// TIA Portal V19 export
ORGANIZATION_BLOCK "CyclicInterrupt"   // OB30, LAD, CyclicInterrupt
{ S7_Optimized_Access := 'TRUE' }
// stored: SetENOAutomatically false
   VAR_INPUT
      Initial_Call : Bool;   // Initial call of this OB
      Event_Count : Int;   // Events discarded
   END_VAR
   VAR_TEMP   // added for the SCL form of the ladder/FBD networks
      _w1 : Bool;
      _w2 : Bool;
   END_VAR
BEGIN

REGION Network 1: CHILLED_P01_SPEED_SP
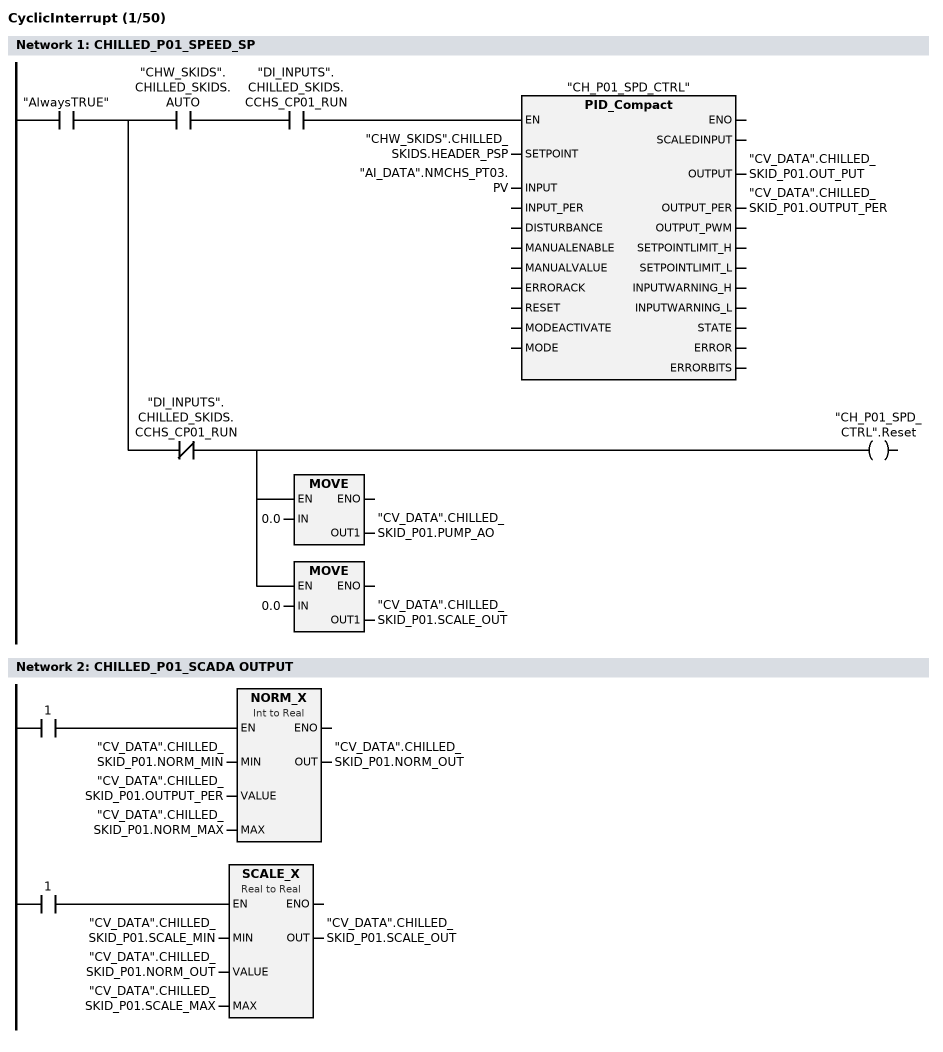
   RUNG wire#powerrail
      Contact( "AlwaysTRUE" )
      wire#w1
      Contact( "CHW_SKIDS".CHILLED_SKIDS.AUTO )
      Contact( "DI_INPUTS".CHILLED_SKIDS.CCHS_CP01_RUN )
      "CH_P01_SPD_CTRL".PID_Compact(Setpoint := "CHW_SKIDS".CHILLED_SKIDS.HEADER_PSP, Input := "AI_DATA".NMCHS_PT03.PV, Input_PER :=, Disturbance :=, ManualEnable :=, ManualValue :=, ErrorAck :=, Reset :=, ModeActivate :=, Mode :=, ScaledInput =>, Output => "CV_DATA".CHILLED_SKID_P01.OUT_PUT, Output_PER => "CV_DATA".CHILLED_SKID_P01.OUTPUT_PER, Output_PWM =>, SetpointLimit_H =>, SetpointLimit_L =>, InputWarning_H =>, InputWarning_L =>, State =>, Error =>, ErrorBits =>)
   END_RUNG
   RUNG wire#w1
      I_Contact( "DI_INPUTS".CHILLED_SKIDS.CCHS_CP01_RUN )
      wire#w2
      Coil( "CH_P01_SPD_CTRL".Reset )
   END_RUNG
   RUNG wire#w2
      Move(in := 0.0, out1 => "CV_DATA".CHILLED_SKID_P01.PUMP_AO)
   END_RUNG
   RUNG wire#w2
      Move(in := 0.0, out1 => "CV_DATA".CHILLED_SKID_P01.SCALE_OUT)
   END_RUNG
   // the same network as SCL:
   #_w1 := "AlwaysTRUE";
   IF "AlwaysTRUE" AND "CHW_SKIDS".CHILLED_SKIDS.AUTO AND "DI_INPUTS".CHILLED_SKIDS.CCHS_CP01_RUN THEN
       "CH_P01_SPD_CTRL"(Setpoint := "CHW_SKIDS".CHILLED_SKIDS.HEADER_PSP,   // PID_Compact
                         Input := "AI_DATA".NMCHS_PT03.PV,
                         Output => "CV_DATA".CHILLED_SKID_P01.OUT_PUT,
                         Output_PER => "CV_DATA".CHILLED_SKID_P01.OUTPUT_PER);
   END_IF;
   "CH_P01_SPD_CTRL".Reset := #_w1 AND NOT "DI_INPUTS".CHILLED_SKIDS.CCHS_CP01_RUN;
   IF "CH_P01_SPD_CTRL".Reset THEN
       "CV_DATA".CHILLED_SKID_P01.PUMP_AO := 0.0;
       "CV_DATA".CHILLED_SKID_P01.SCALE_OUT := 0.0;
   END_IF;
END_REGION

REGION Network 2: CHILLED_P01_SCADA OUTPUT
   RUNG wire#powerrail
      Contact( 1 )
      { S7_Templates := "[SrcType := Int, DestType := Real]" } Normalize(min := "CV_DATA".CHILLED_SKID_P01.NORM_MIN, value := "CV_DATA".CHILLED_SKID_P01.OUTPUT_PER, max := "CV_DATA".CHILLED_SKID_P01.NORM_MAX, out => "CV_DATA".CHILLED_SKID_P01.NORM_OUT)
   END_RUNG
   RUNG wire#powerrail
      Contact( 1 )
      { S7_Templates := "[SrcType := Real, DestType := Real]" } Scale(min := "CV_DATA".CHILLED_SKID_P01.SCALE_MIN, value := "CV_DATA".CHILLED_SKID_P01.NORM_OUT, max := "CV_DATA".CHILLED_SKID_P01.SCALE_MAX, out => "CV_DATA".CHILLED_SKID_P01.SCALE_OUT)
   END_RUNG
   // the same network as SCL:
   IF 1 THEN
       "CV_DATA".CHILLED_SKID_P01.NORM_OUT := NORM_X(MIN := "CV_DATA".CHILLED_SKID_P01.NORM_MIN, VALUE := "CV_DATA".CHILLED_SKID_P01.OUTPUT_PER, MAX := "CV_DATA".CHILLED_SKID_P01.NORM_MAX);
       "CV_DATA".CHILLED_SKID_P01.SCALE_OUT := SCALE_X(MIN := "CV_DATA".CHILLED_SKID_P01.SCALE_MIN, VALUE := "CV_DATA".CHILLED_SKID_P01.NORM_OUT, MAX := "CV_DATA".CHILLED_SKID_P01.SCALE_MAX);
   END_IF;
END_REGION

REGION Network 3: CHILLED_P01_MANUAL OUTPUT
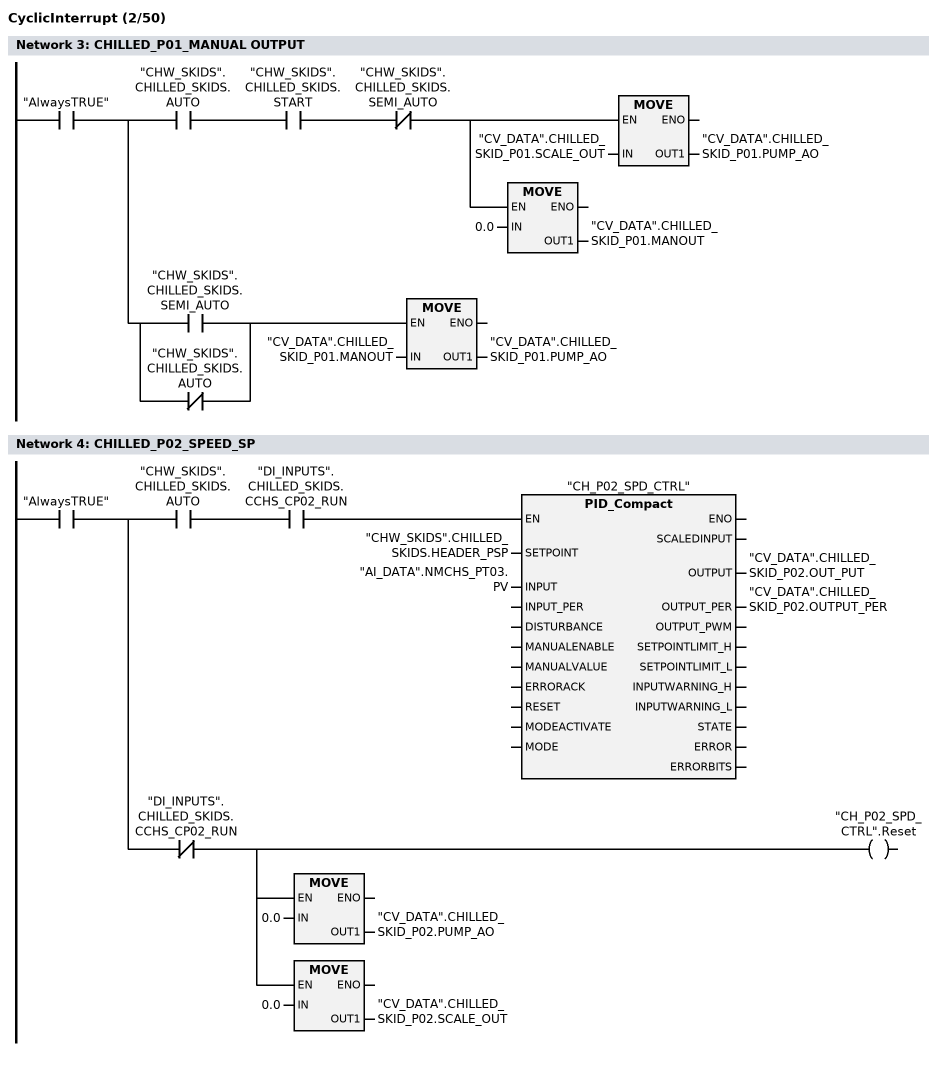
   RUNG wire#powerrail
      Contact( "AlwaysTRUE" )
      wire#w1
      Contact( "CHW_SKIDS".CHILLED_SKIDS.AUTO )
      Contact( "CHW_SKIDS".CHILLED_SKIDS.START )
      I_Contact( "CHW_SKIDS".CHILLED_SKIDS.SEMI_AUTO )
      wire#w2
      Move(in := "CV_DATA".CHILLED_SKID_P01.SCALE_OUT, out1 => "CV_DATA".CHILLED_SKID_P01.PUMP_AO)
   END_RUNG
   RUNG wire#w2
      Move(in := 0.0, out1 => "CV_DATA".CHILLED_SKID_P01.MANOUT)
   END_RUNG
   RUNG wire#w1
      Contact( "CHW_SKIDS".CHILLED_SKIDS.SEMI_AUTO )
      wire#w3
      Move(in := "CV_DATA".CHILLED_SKID_P01.MANOUT, out1 => "CV_DATA".CHILLED_SKID_P01.PUMP_AO)
   END_RUNG
   RUNG wire#w1
      I_Contact( "CHW_SKIDS".CHILLED_SKIDS.AUTO )
   END_RUNG wire#w3
   // the same network as SCL:
   IF "AlwaysTRUE" AND "CHW_SKIDS".CHILLED_SKIDS.AUTO AND "CHW_SKIDS".CHILLED_SKIDS.START AND NOT "CHW_SKIDS".CHILLED_SKIDS.SEMI_AUTO THEN
       "CV_DATA".CHILLED_SKID_P01.PUMP_AO := "CV_DATA".CHILLED_SKID_P01.SCALE_OUT;
       "CV_DATA".CHILLED_SKID_P01.MANOUT := 0.0;
   END_IF;
   IF "AlwaysTRUE" AND ("CHW_SKIDS".CHILLED_SKIDS.SEMI_AUTO OR NOT "CHW_SKIDS".CHILLED_SKIDS.AUTO) THEN
       "CV_DATA".CHILLED_SKID_P01.PUMP_AO := "CV_DATA".CHILLED_SKID_P01.MANOUT;
   END_IF;
END_REGION

REGION Network 4: CHILLED_P02_SPEED_SP
   RUNG wire#powerrail
      Contact( "AlwaysTRUE" )
      wire#w1
      Contact( "CHW_SKIDS".CHILLED_SKIDS.AUTO )
      Contact( "DI_INPUTS".CHILLED_SKIDS.CCHS_CP02_RUN )
      "CH_P02_SPD_CTRL".PID_Compact(Setpoint := "CHW_SKIDS".CHILLED_SKIDS.HEADER_PSP, Input := "AI_DATA".NMCHS_PT03.PV, Input_PER :=, Disturbance :=, ManualEnable :=, ManualValue :=, ErrorAck :=, Reset :=, ModeActivate :=, Mode :=, ScaledInput =>, Output => "CV_DATA".CHILLED_SKID_P02.OUT_PUT, Output_PER => "CV_DATA".CHILLED_SKID_P02.OUTPUT_PER, Output_PWM =>, SetpointLimit_H =>, SetpointLimit_L =>, InputWarning_H =>, InputWarning_L =>, State =>, Error =>, ErrorBits =>)
   END_RUNG
   RUNG wire#w1
      I_Contact( "DI_INPUTS".CHILLED_SKIDS.CCHS_CP02_RUN )
      wire#w2
      Coil( "CH_P02_SPD_CTRL".Reset )
   END_RUNG
   RUNG wire#w2
      Move(in := 0.0, out1 => "CV_DATA".CHILLED_SKID_P02.PUMP_AO)
   END_RUNG
   RUNG wire#w2
      Move(in := 0.0, out1 => "CV_DATA".CHILLED_SKID_P02.SCALE_OUT)
   END_RUNG
   // the same network as SCL:
   #_w1 := "AlwaysTRUE";
   IF "AlwaysTRUE" AND "CHW_SKIDS".CHILLED_SKIDS.AUTO AND "DI_INPUTS".CHILLED_SKIDS.CCHS_CP02_RUN THEN
       "CH_P02_SPD_CTRL"(Setpoint := "CHW_SKIDS".CHILLED_SKIDS.HEADER_PSP,   // PID_Compact
                         Input := "AI_DATA".NMCHS_PT03.PV,
                         Output => "CV_DATA".CHILLED_SKID_P02.OUT_PUT,
                         Output_PER => "CV_DATA".CHILLED_SKID_P02.OUTPUT_PER);
   END_IF;
   "CH_P02_SPD_CTRL".Reset := #_w1 AND NOT "DI_INPUTS".CHILLED_SKIDS.CCHS_CP02_RUN;
   IF "CH_P02_SPD_CTRL".Reset THEN
       "CV_DATA".CHILLED_SKID_P02.PUMP_AO := 0.0;
       "CV_DATA".CHILLED_SKID_P02.SCALE_OUT := 0.0;
   END_IF;
END_REGION

REGION Network 5: CHILLED_P02_SCADA OUTPUT
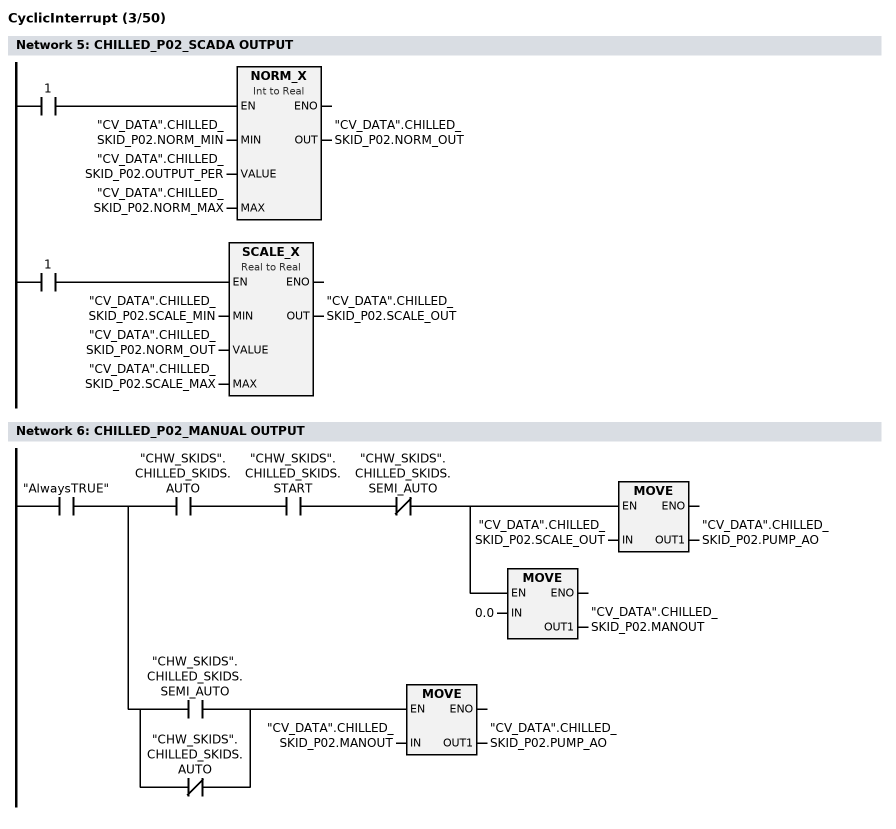
   RUNG wire#powerrail
      Contact( 1 )
      { S7_Templates := "[SrcType := Int, DestType := Real]" } Normalize(min := "CV_DATA".CHILLED_SKID_P02.NORM_MIN, value := "CV_DATA".CHILLED_SKID_P02.OUTPUT_PER, max := "CV_DATA".CHILLED_SKID_P02.NORM_MAX, out => "CV_DATA".CHILLED_SKID_P02.NORM_OUT)
   END_RUNG
   RUNG wire#powerrail
      Contact( 1 )
      { S7_Templates := "[SrcType := Real, DestType := Real]" } Scale(min := "CV_DATA".CHILLED_SKID_P02.SCALE_MIN, value := "CV_DATA".CHILLED_SKID_P02.NORM_OUT, max := "CV_DATA".CHILLED_SKID_P02.SCALE_MAX, out => "CV_DATA".CHILLED_SKID_P02.SCALE_OUT)
   END_RUNG
   // the same network as SCL:
   IF 1 THEN
       "CV_DATA".CHILLED_SKID_P02.NORM_OUT := NORM_X(MIN := "CV_DATA".CHILLED_SKID_P02.NORM_MIN, VALUE := "CV_DATA".CHILLED_SKID_P02.OUTPUT_PER, MAX := "CV_DATA".CHILLED_SKID_P02.NORM_MAX);
       "CV_DATA".CHILLED_SKID_P02.SCALE_OUT := SCALE_X(MIN := "CV_DATA".CHILLED_SKID_P02.SCALE_MIN, VALUE := "CV_DATA".CHILLED_SKID_P02.NORM_OUT, MAX := "CV_DATA".CHILLED_SKID_P02.SCALE_MAX);
   END_IF;
END_REGION

REGION Network 6: CHILLED_P02_MANUAL OUTPUT
   RUNG wire#powerrail
      Contact( "AlwaysTRUE" )
      wire#w1
      Contact( "CHW_SKIDS".CHILLED_SKIDS.AUTO )
      Contact( "CHW_SKIDS".CHILLED_SKIDS.START )
      I_Contact( "CHW_SKIDS".CHILLED_SKIDS.SEMI_AUTO )
      wire#w2
      Move(in := "CV_DATA".CHILLED_SKID_P02.SCALE_OUT, out1 => "CV_DATA".CHILLED_SKID_P02.PUMP_AO)
   END_RUNG
   RUNG wire#w2
      Move(in := 0.0, out1 => "CV_DATA".CHILLED_SKID_P02.MANOUT)
   END_RUNG
   RUNG wire#w1
      Contact( "CHW_SKIDS".CHILLED_SKIDS.SEMI_AUTO )
      wire#w3
      Move(in := "CV_DATA".CHILLED_SKID_P02.MANOUT, out1 => "CV_DATA".CHILLED_SKID_P02.PUMP_AO)
   END_RUNG
   RUNG wire#w1
      I_Contact( "CHW_SKIDS".CHILLED_SKIDS.AUTO )
   END_RUNG wire#w3
   // the same network as SCL:
   IF "AlwaysTRUE" AND "CHW_SKIDS".CHILLED_SKIDS.AUTO AND "CHW_SKIDS".CHILLED_SKIDS.START AND NOT "CHW_SKIDS".CHILLED_SKIDS.SEMI_AUTO THEN
       "CV_DATA".CHILLED_SKID_P02.PUMP_AO := "CV_DATA".CHILLED_SKID_P02.SCALE_OUT;
       "CV_DATA".CHILLED_SKID_P02.MANOUT := 0.0;
   END_IF;
   IF "AlwaysTRUE" AND ("CHW_SKIDS".CHILLED_SKIDS.SEMI_AUTO OR NOT "CHW_SKIDS".CHILLED_SKIDS.AUTO) THEN
       "CV_DATA".CHILLED_SKID_P02.PUMP_AO := "CV_DATA".CHILLED_SKID_P02.MANOUT;
   END_IF;
END_REGION

REGION Network 7: CHILLED_P03_SPEED_SP
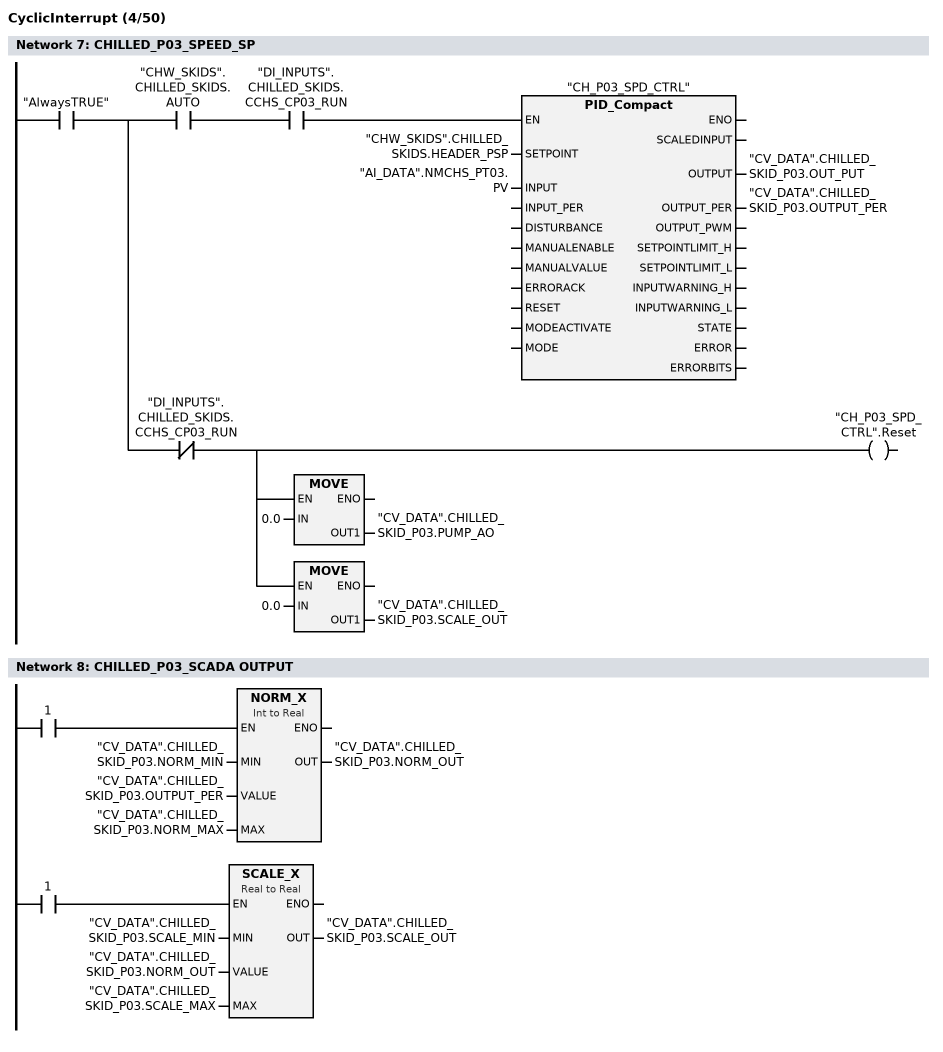
   RUNG wire#powerrail
      Contact( "AlwaysTRUE" )
      wire#w1
      Contact( "CHW_SKIDS".CHILLED_SKIDS.AUTO )
      Contact( "DI_INPUTS".CHILLED_SKIDS.CCHS_CP03_RUN )
      "CH_P03_SPD_CTRL".PID_Compact(Setpoint := "CHW_SKIDS".CHILLED_SKIDS.HEADER_PSP, Input := "AI_DATA".NMCHS_PT03.PV, Input_PER :=, Disturbance :=, ManualEnable :=, ManualValue :=, ErrorAck :=, Reset :=, ModeActivate :=, Mode :=, ScaledInput =>, Output => "CV_DATA".CHILLED_SKID_P03.OUT_PUT, Output_PER => "CV_DATA".CHILLED_SKID_P03.OUTPUT_PER, Output_PWM =>, SetpointLimit_H =>, SetpointLimit_L =>, InputWarning_H =>, InputWarning_L =>, State =>, Error =>, ErrorBits =>)
   END_RUNG
   RUNG wire#w1
      I_Contact( "DI_INPUTS".CHILLED_SKIDS.CCHS_CP03_RUN )
      wire#w2
      Coil( "CH_P03_SPD_CTRL".Reset )
   END_RUNG
   RUNG wire#w2
      Move(in := 0.0, out1 => "CV_DATA".CHILLED_SKID_P03.PUMP_AO)
   END_RUNG
   RUNG wire#w2
      Move(in := 0.0, out1 => "CV_DATA".CHILLED_SKID_P03.SCALE_OUT)
   END_RUNG
   // the same network as SCL:
   #_w1 := "AlwaysTRUE";
   IF "AlwaysTRUE" AND "CHW_SKIDS".CHILLED_SKIDS.AUTO AND "DI_INPUTS".CHILLED_SKIDS.CCHS_CP03_RUN THEN
       "CH_P03_SPD_CTRL"(Setpoint := "CHW_SKIDS".CHILLED_SKIDS.HEADER_PSP,   // PID_Compact
                         Input := "AI_DATA".NMCHS_PT03.PV,
                         Output => "CV_DATA".CHILLED_SKID_P03.OUT_PUT,
                         Output_PER => "CV_DATA".CHILLED_SKID_P03.OUTPUT_PER);
   END_IF;
   "CH_P03_SPD_CTRL".Reset := #_w1 AND NOT "DI_INPUTS".CHILLED_SKIDS.CCHS_CP03_RUN;
   IF "CH_P03_SPD_CTRL".Reset THEN
       "CV_DATA".CHILLED_SKID_P03.PUMP_AO := 0.0;
       "CV_DATA".CHILLED_SKID_P03.SCALE_OUT := 0.0;
   END_IF;
END_REGION

REGION Network 8: CHILLED_P03_SCADA OUTPUT
   RUNG wire#powerrail
      Contact( 1 )
      { S7_Templates := "[SrcType := Int, DestType := Real]" } Normalize(min := "CV_DATA".CHILLED_SKID_P03.NORM_MIN, value := "CV_DATA".CHILLED_SKID_P03.OUTPUT_PER, max := "CV_DATA".CHILLED_SKID_P03.NORM_MAX, out => "CV_DATA".CHILLED_SKID_P03.NORM_OUT)
   END_RUNG
   RUNG wire#powerrail
      Contact( 1 )
      { S7_Templates := "[SrcType := Real, DestType := Real]" } Scale(min := "CV_DATA".CHILLED_SKID_P03.SCALE_MIN, value := "CV_DATA".CHILLED_SKID_P03.NORM_OUT, max := "CV_DATA".CHILLED_SKID_P03.SCALE_MAX, out => "CV_DATA".CHILLED_SKID_P03.SCALE_OUT)
   END_RUNG
   // the same network as SCL:
   IF 1 THEN
       "CV_DATA".CHILLED_SKID_P03.NORM_OUT := NORM_X(MIN := "CV_DATA".CHILLED_SKID_P03.NORM_MIN, VALUE := "CV_DATA".CHILLED_SKID_P03.OUTPUT_PER, MAX := "CV_DATA".CHILLED_SKID_P03.NORM_MAX);
       "CV_DATA".CHILLED_SKID_P03.SCALE_OUT := SCALE_X(MIN := "CV_DATA".CHILLED_SKID_P03.SCALE_MIN, VALUE := "CV_DATA".CHILLED_SKID_P03.NORM_OUT, MAX := "CV_DATA".CHILLED_SKID_P03.SCALE_MAX);
   END_IF;
END_REGION

REGION Network 9: CHILLED_P03_MANUAL OUTPUT
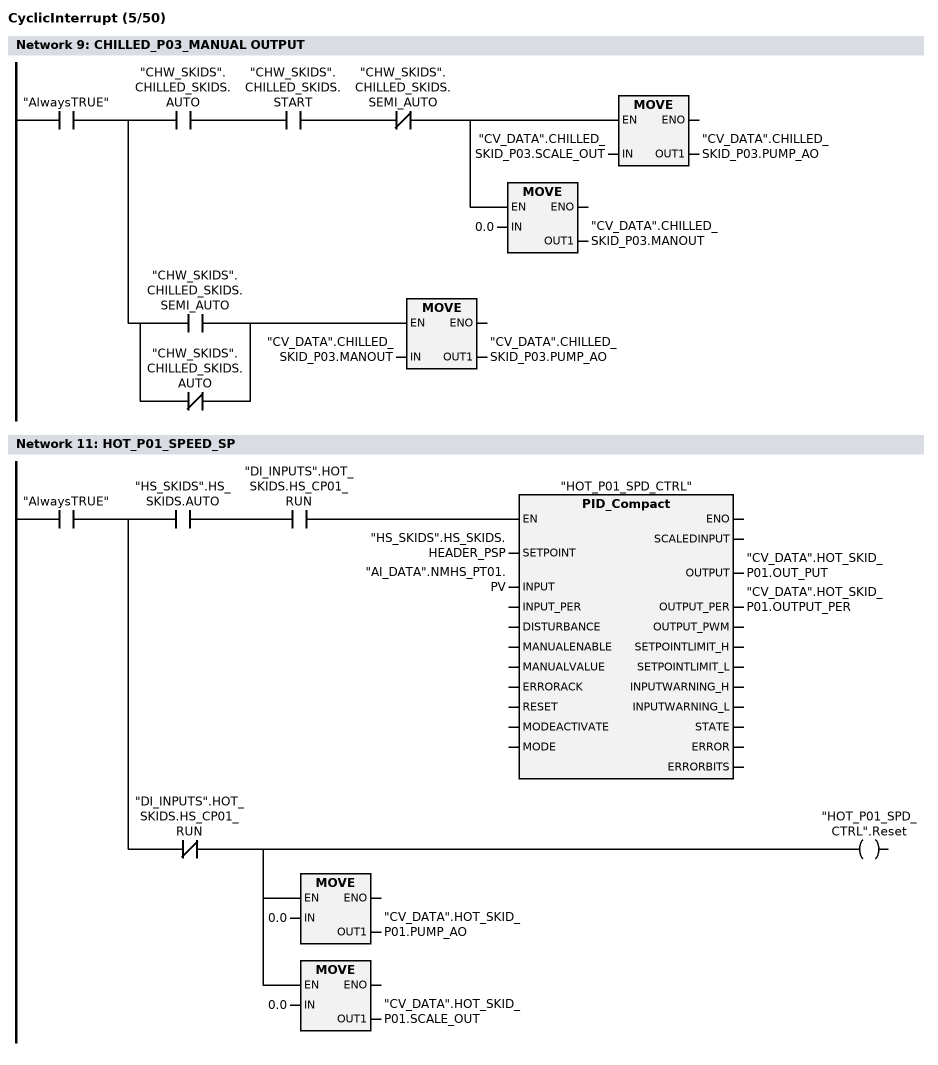
   RUNG wire#powerrail
      Contact( "AlwaysTRUE" )
      wire#w1
      Contact( "CHW_SKIDS".CHILLED_SKIDS.AUTO )
      Contact( "CHW_SKIDS".CHILLED_SKIDS.START )
      I_Contact( "CHW_SKIDS".CHILLED_SKIDS.SEMI_AUTO )
      wire#w2
      Move(in := "CV_DATA".CHILLED_SKID_P03.SCALE_OUT, out1 => "CV_DATA".CHILLED_SKID_P03.PUMP_AO)
   END_RUNG
   RUNG wire#w2
      Move(in := 0.0, out1 => "CV_DATA".CHILLED_SKID_P03.MANOUT)
   END_RUNG
   RUNG wire#w1
      Contact( "CHW_SKIDS".CHILLED_SKIDS.SEMI_AUTO )
      wire#w3
      Move(in := "CV_DATA".CHILLED_SKID_P03.MANOUT, out1 => "CV_DATA".CHILLED_SKID_P03.PUMP_AO)
   END_RUNG
   RUNG wire#w1
      I_Contact( "CHW_SKIDS".CHILLED_SKIDS.AUTO )
   END_RUNG wire#w3
   // the same network as SCL:
   IF "AlwaysTRUE" AND "CHW_SKIDS".CHILLED_SKIDS.AUTO AND "CHW_SKIDS".CHILLED_SKIDS.START AND NOT "CHW_SKIDS".CHILLED_SKIDS.SEMI_AUTO THEN
       "CV_DATA".CHILLED_SKID_P03.PUMP_AO := "CV_DATA".CHILLED_SKID_P03.SCALE_OUT;
       "CV_DATA".CHILLED_SKID_P03.MANOUT := 0.0;
   END_IF;
   IF "AlwaysTRUE" AND ("CHW_SKIDS".CHILLED_SKIDS.SEMI_AUTO OR NOT "CHW_SKIDS".CHILLED_SKIDS.AUTO) THEN
       "CV_DATA".CHILLED_SKID_P03.PUMP_AO := "CV_DATA".CHILLED_SKID_P03.MANOUT;
   END_IF;
END_REGION

REGION Network 11: HOT_P01_SPEED_SP
   RUNG wire#powerrail
      Contact( "AlwaysTRUE" )
      wire#w1
      Contact( "HS_SKIDS".HS_SKIDS.AUTO )
      Contact( "DI_INPUTS".HOT_SKIDS.HS_CP01_RUN )
      "HOT_P01_SPD_CTRL".PID_Compact(Setpoint := "HS_SKIDS".HS_SKIDS.HEADER_PSP, Input := "AI_DATA".NMHS_PT01.PV, Input_PER :=, Disturbance :=, ManualEnable :=, ManualValue :=, ErrorAck :=, Reset :=, ModeActivate :=, Mode :=, ScaledInput =>, Output => "CV_DATA".HOT_SKID_P01.OUT_PUT, Output_PER => "CV_DATA".HOT_SKID_P01.OUTPUT_PER, Output_PWM =>, SetpointLimit_H =>, SetpointLimit_L =>, InputWarning_H =>, InputWarning_L =>, State =>, Error =>, ErrorBits =>)
   END_RUNG
   RUNG wire#w1
      I_Contact( "DI_INPUTS".HOT_SKIDS.HS_CP01_RUN )
      wire#w2
      Coil( "HOT_P01_SPD_CTRL".Reset )
   END_RUNG
   RUNG wire#w2
      Move(in := 0.0, out1 => "CV_DATA".HOT_SKID_P01.PUMP_AO)
   END_RUNG
   RUNG wire#w2
      Move(in := 0.0, out1 => "CV_DATA".HOT_SKID_P01.SCALE_OUT)
   END_RUNG
   // the same network as SCL:
   #_w1 := "AlwaysTRUE";
   IF "AlwaysTRUE" AND "HS_SKIDS".HS_SKIDS.AUTO AND "DI_INPUTS".HOT_SKIDS.HS_CP01_RUN THEN
       "HOT_P01_SPD_CTRL"(Setpoint := "HS_SKIDS".HS_SKIDS.HEADER_PSP,   // PID_Compact
                          Input := "AI_DATA".NMHS_PT01.PV,
                          Output => "CV_DATA".HOT_SKID_P01.OUT_PUT,
                          Output_PER => "CV_DATA".HOT_SKID_P01.OUTPUT_PER);
   END_IF;
   "HOT_P01_SPD_CTRL".Reset := #_w1 AND NOT "DI_INPUTS".HOT_SKIDS.HS_CP01_RUN;
   IF "HOT_P01_SPD_CTRL".Reset THEN
       "CV_DATA".HOT_SKID_P01.PUMP_AO := 0.0;
       "CV_DATA".HOT_SKID_P01.SCALE_OUT := 0.0;
   END_IF;
END_REGION

REGION Network 12: HOT_P01_SCADA OUTPUT
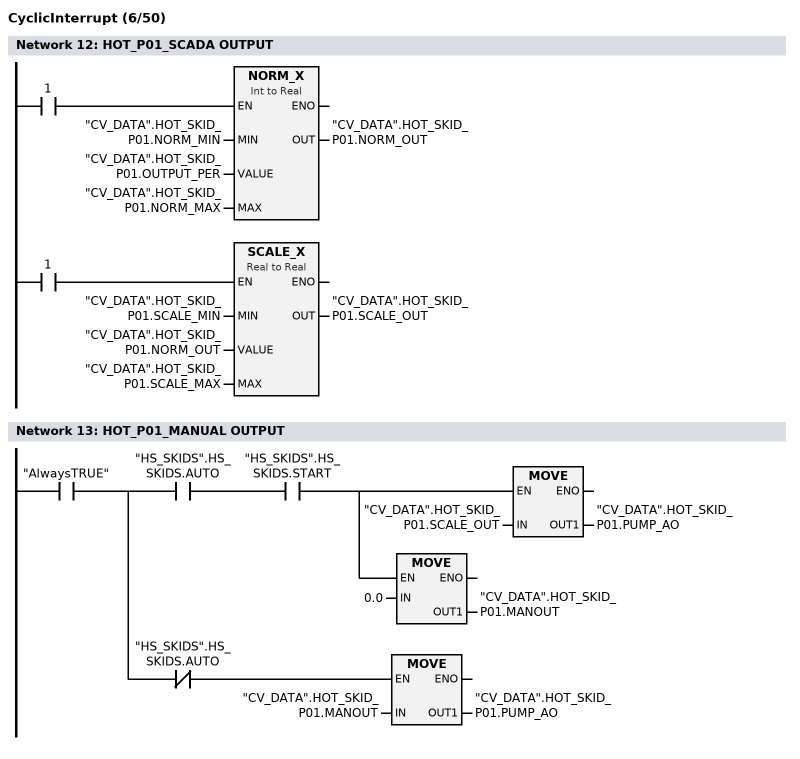
   RUNG wire#powerrail
      Contact( 1 )
      { S7_Templates := "[SrcType := Int, DestType := Real]" } Normalize(min := "CV_DATA".HOT_SKID_P01.NORM_MIN, value := "CV_DATA".HOT_SKID_P01.OUTPUT_PER, max := "CV_DATA".HOT_SKID_P01.NORM_MAX, out => "CV_DATA".HOT_SKID_P01.NORM_OUT)
   END_RUNG
   RUNG wire#powerrail
      Contact( 1 )
      { S7_Templates := "[SrcType := Real, DestType := Real]" } Scale(min := "CV_DATA".HOT_SKID_P01.SCALE_MIN, value := "CV_DATA".HOT_SKID_P01.NORM_OUT, max := "CV_DATA".HOT_SKID_P01.SCALE_MAX, out => "CV_DATA".HOT_SKID_P01.SCALE_OUT)
   END_RUNG
   // the same network as SCL:
   IF 1 THEN
       "CV_DATA".HOT_SKID_P01.NORM_OUT := NORM_X(MIN := "CV_DATA".HOT_SKID_P01.NORM_MIN, VALUE := "CV_DATA".HOT_SKID_P01.OUTPUT_PER, MAX := "CV_DATA".HOT_SKID_P01.NORM_MAX);
       "CV_DATA".HOT_SKID_P01.SCALE_OUT := SCALE_X(MIN := "CV_DATA".HOT_SKID_P01.SCALE_MIN, VALUE := "CV_DATA".HOT_SKID_P01.NORM_OUT, MAX := "CV_DATA".HOT_SKID_P01.SCALE_MAX);
   END_IF;
END_REGION

REGION Network 13: HOT_P01_MANUAL OUTPUT
   RUNG wire#powerrail
      Contact( "AlwaysTRUE" )
      wire#w1
      Contact( "HS_SKIDS".HS_SKIDS.AUTO )
      Contact( "HS_SKIDS".HS_SKIDS.START )
      wire#w2
      Move(in := "CV_DATA".HOT_SKID_P01.SCALE_OUT, out1 => "CV_DATA".HOT_SKID_P01.PUMP_AO)
   END_RUNG
   RUNG wire#w2
      Move(in := 0.0, out1 => "CV_DATA".HOT_SKID_P01.MANOUT)
   END_RUNG
   RUNG wire#w1
      I_Contact( "HS_SKIDS".HS_SKIDS.AUTO )
      Move(in := "CV_DATA".HOT_SKID_P01.MANOUT, out1 => "CV_DATA".HOT_SKID_P01.PUMP_AO)
   END_RUNG
   // the same network as SCL:
   IF "AlwaysTRUE" AND "HS_SKIDS".HS_SKIDS.AUTO AND "HS_SKIDS".HS_SKIDS.START THEN
       "CV_DATA".HOT_SKID_P01.PUMP_AO := "CV_DATA".HOT_SKID_P01.SCALE_OUT;
       "CV_DATA".HOT_SKID_P01.MANOUT := 0.0;
   END_IF;
   IF "AlwaysTRUE" AND NOT "HS_SKIDS".HS_SKIDS.AUTO THEN
       "CV_DATA".HOT_SKID_P01.PUMP_AO := "CV_DATA".HOT_SKID_P01.MANOUT;
   END_IF;
END_REGION

REGION Network 14: HOT_P02_SPEED_SP
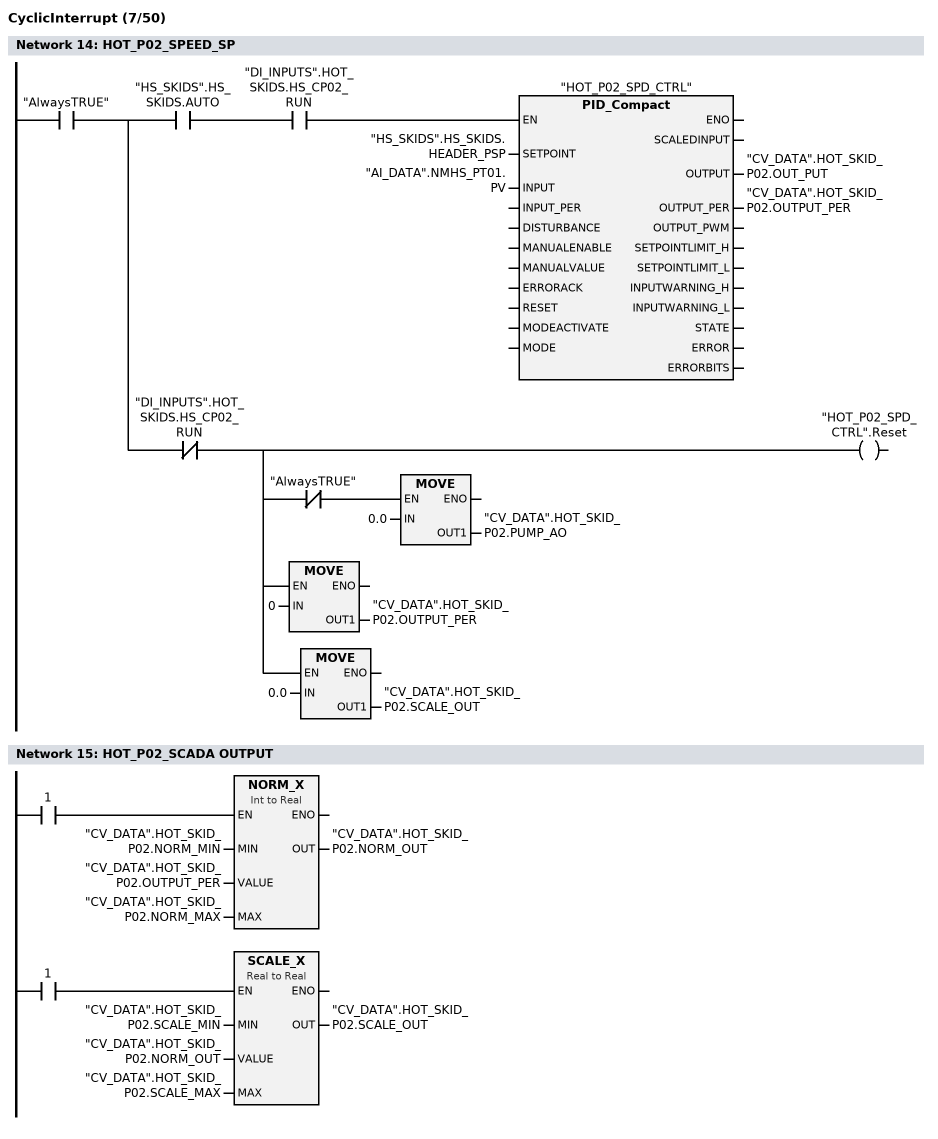
   RUNG wire#powerrail
      Contact( "AlwaysTRUE" )
      wire#w1
      Contact( "HS_SKIDS".HS_SKIDS.AUTO )
      Contact( "DI_INPUTS".HOT_SKIDS.HS_CP02_RUN )
      "HOT_P02_SPD_CTRL".PID_Compact(Setpoint := "HS_SKIDS".HS_SKIDS.HEADER_PSP, Input := "AI_DATA".NMHS_PT01.PV, Input_PER :=, Disturbance :=, ManualEnable :=, ManualValue :=, ErrorAck :=, Reset :=, ModeActivate :=, Mode :=, ScaledInput =>, Output => "CV_DATA".HOT_SKID_P02.OUT_PUT, Output_PER => "CV_DATA".HOT_SKID_P02.OUTPUT_PER, Output_PWM =>, SetpointLimit_H =>, SetpointLimit_L =>, InputWarning_H =>, InputWarning_L =>, State =>, Error =>, ErrorBits =>)
   END_RUNG
   RUNG wire#w1
      I_Contact( "DI_INPUTS".HOT_SKIDS.HS_CP02_RUN )
      wire#w2
      Coil( "HOT_P02_SPD_CTRL".Reset )
   END_RUNG
   RUNG wire#w2
      I_Contact( "AlwaysTRUE" )
      Move(in := 0.0, out1 => "CV_DATA".HOT_SKID_P02.PUMP_AO)
   END_RUNG
   RUNG wire#w2
      Move(in := 0, out1 => "CV_DATA".HOT_SKID_P02.OUTPUT_PER)
   END_RUNG
   RUNG wire#w2
      Move(in := 0.0, out1 => "CV_DATA".HOT_SKID_P02.SCALE_OUT)
   END_RUNG
   // the same network as SCL:
   #_w1 := "AlwaysTRUE";
   IF "AlwaysTRUE" AND "HS_SKIDS".HS_SKIDS.AUTO AND "DI_INPUTS".HOT_SKIDS.HS_CP02_RUN THEN
       "HOT_P02_SPD_CTRL"(Setpoint := "HS_SKIDS".HS_SKIDS.HEADER_PSP,   // PID_Compact
                          Input := "AI_DATA".NMHS_PT01.PV,
                          Output => "CV_DATA".HOT_SKID_P02.OUT_PUT,
                          Output_PER => "CV_DATA".HOT_SKID_P02.OUTPUT_PER);
   END_IF;
   "HOT_P02_SPD_CTRL".Reset := #_w1 AND NOT "DI_INPUTS".HOT_SKIDS.HS_CP02_RUN;
   IF "HOT_P02_SPD_CTRL".Reset AND NOT "AlwaysTRUE" THEN "CV_DATA".HOT_SKID_P02.PUMP_AO := 0.0; END_IF;
   IF "HOT_P02_SPD_CTRL".Reset THEN
       "CV_DATA".HOT_SKID_P02.OUTPUT_PER := 0;
       "CV_DATA".HOT_SKID_P02.SCALE_OUT := 0.0;
   END_IF;
END_REGION

REGION Network 15: HOT_P02_SCADA OUTPUT
   RUNG wire#powerrail
      Contact( 1 )
      { S7_Templates := "[SrcType := Int, DestType := Real]" } Normalize(min := "CV_DATA".HOT_SKID_P02.NORM_MIN, value := "CV_DATA".HOT_SKID_P02.OUTPUT_PER, max := "CV_DATA".HOT_SKID_P02.NORM_MAX, out => "CV_DATA".HOT_SKID_P02.NORM_OUT)
   END_RUNG
   RUNG wire#powerrail
      Contact( 1 )
      { S7_Templates := "[SrcType := Real, DestType := Real]" } Scale(min := "CV_DATA".HOT_SKID_P02.SCALE_MIN, value := "CV_DATA".HOT_SKID_P02.NORM_OUT, max := "CV_DATA".HOT_SKID_P02.SCALE_MAX, out => "CV_DATA".HOT_SKID_P02.SCALE_OUT)
   END_RUNG
   // the same network as SCL:
   IF 1 THEN
       "CV_DATA".HOT_SKID_P02.NORM_OUT := NORM_X(MIN := "CV_DATA".HOT_SKID_P02.NORM_MIN, VALUE := "CV_DATA".HOT_SKID_P02.OUTPUT_PER, MAX := "CV_DATA".HOT_SKID_P02.NORM_MAX);
       "CV_DATA".HOT_SKID_P02.SCALE_OUT := SCALE_X(MIN := "CV_DATA".HOT_SKID_P02.SCALE_MIN, VALUE := "CV_DATA".HOT_SKID_P02.NORM_OUT, MAX := "CV_DATA".HOT_SKID_P02.SCALE_MAX);
   END_IF;
END_REGION

REGION Network 16: HOT_P02_MANUAL OUTPUT
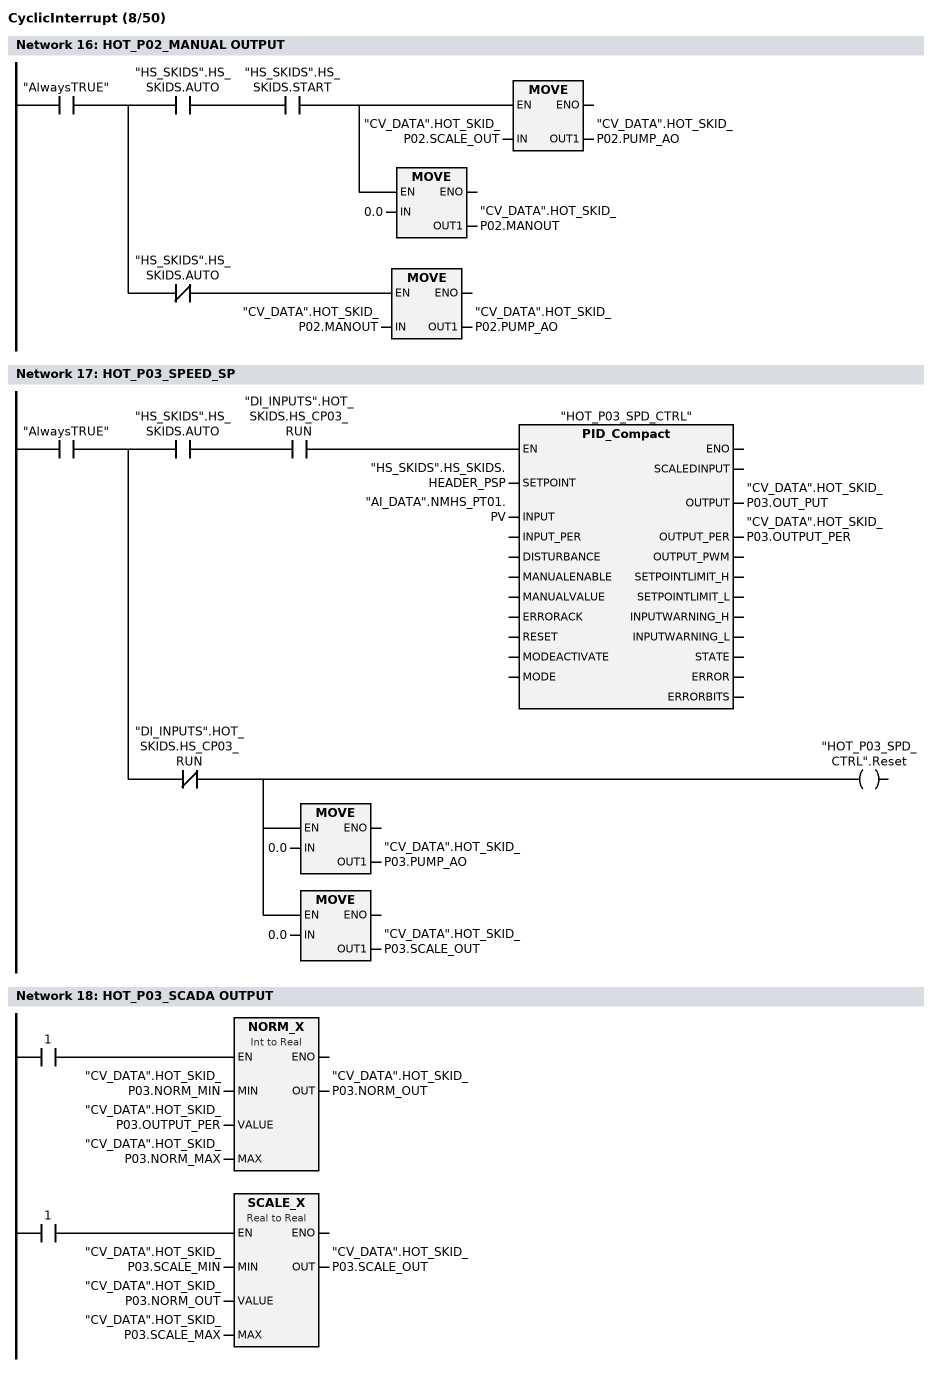
   RUNG wire#powerrail
      Contact( "AlwaysTRUE" )
      wire#w1
      Contact( "HS_SKIDS".HS_SKIDS.AUTO )
      Contact( "HS_SKIDS".HS_SKIDS.START )
      wire#w2
      Move(in := "CV_DATA".HOT_SKID_P02.SCALE_OUT, out1 => "CV_DATA".HOT_SKID_P02.PUMP_AO)
   END_RUNG
   RUNG wire#w2
      Move(in := 0.0, out1 => "CV_DATA".HOT_SKID_P02.MANOUT)
   END_RUNG
   RUNG wire#w1
      I_Contact( "HS_SKIDS".HS_SKIDS.AUTO )
      Move(in := "CV_DATA".HOT_SKID_P02.MANOUT, out1 => "CV_DATA".HOT_SKID_P02.PUMP_AO)
   END_RUNG
   // the same network as SCL:
   IF "AlwaysTRUE" AND "HS_SKIDS".HS_SKIDS.AUTO AND "HS_SKIDS".HS_SKIDS.START THEN
       "CV_DATA".HOT_SKID_P02.PUMP_AO := "CV_DATA".HOT_SKID_P02.SCALE_OUT;
       "CV_DATA".HOT_SKID_P02.MANOUT := 0.0;
   END_IF;
   IF "AlwaysTRUE" AND NOT "HS_SKIDS".HS_SKIDS.AUTO THEN
       "CV_DATA".HOT_SKID_P02.PUMP_AO := "CV_DATA".HOT_SKID_P02.MANOUT;
   END_IF;
END_REGION

REGION Network 17: HOT_P03_SPEED_SP
   RUNG wire#powerrail
      Contact( "AlwaysTRUE" )
      wire#w1
      Contact( "HS_SKIDS".HS_SKIDS.AUTO )
      Contact( "DI_INPUTS".HOT_SKIDS.HS_CP03_RUN )
      "HOT_P03_SPD_CTRL".PID_Compact(Setpoint := "HS_SKIDS".HS_SKIDS.HEADER_PSP, Input := "AI_DATA".NMHS_PT01.PV, Input_PER :=, Disturbance :=, ManualEnable :=, ManualValue :=, ErrorAck :=, Reset :=, ModeActivate :=, Mode :=, ScaledInput =>, Output => "CV_DATA".HOT_SKID_P03.OUT_PUT, Output_PER => "CV_DATA".HOT_SKID_P03.OUTPUT_PER, Output_PWM =>, SetpointLimit_H =>, SetpointLimit_L =>, InputWarning_H =>, InputWarning_L =>, State =>, Error =>, ErrorBits =>)
   END_RUNG
   RUNG wire#w1
      I_Contact( "DI_INPUTS".HOT_SKIDS.HS_CP03_RUN )
      wire#w2
      Coil( "HOT_P03_SPD_CTRL".Reset )
   END_RUNG
   RUNG wire#w2
      Move(in := 0.0, out1 => "CV_DATA".HOT_SKID_P03.PUMP_AO)
   END_RUNG
   RUNG wire#w2
      Move(in := 0.0, out1 => "CV_DATA".HOT_SKID_P03.SCALE_OUT)
   END_RUNG
   // the same network as SCL:
   #_w1 := "AlwaysTRUE";
   IF "AlwaysTRUE" AND "HS_SKIDS".HS_SKIDS.AUTO AND "DI_INPUTS".HOT_SKIDS.HS_CP03_RUN THEN
       "HOT_P03_SPD_CTRL"(Setpoint := "HS_SKIDS".HS_SKIDS.HEADER_PSP,   // PID_Compact
                          Input := "AI_DATA".NMHS_PT01.PV,
                          Output => "CV_DATA".HOT_SKID_P03.OUT_PUT,
                          Output_PER => "CV_DATA".HOT_SKID_P03.OUTPUT_PER);
   END_IF;
   "HOT_P03_SPD_CTRL".Reset := #_w1 AND NOT "DI_INPUTS".HOT_SKIDS.HS_CP03_RUN;
   IF "HOT_P03_SPD_CTRL".Reset THEN
       "CV_DATA".HOT_SKID_P03.PUMP_AO := 0.0;
       "CV_DATA".HOT_SKID_P03.SCALE_OUT := 0.0;
   END_IF;
END_REGION

REGION Network 18: HOT_P03_SCADA OUTPUT
   RUNG wire#powerrail
      Contact( 1 )
      { S7_Templates := "[SrcType := Int, DestType := Real]" } Normalize(min := "CV_DATA".HOT_SKID_P03.NORM_MIN, value := "CV_DATA".HOT_SKID_P03.OUTPUT_PER, max := "CV_DATA".HOT_SKID_P03.NORM_MAX, out => "CV_DATA".HOT_SKID_P03.NORM_OUT)
   END_RUNG
   RUNG wire#powerrail
      Contact( 1 )
      { S7_Templates := "[SrcType := Real, DestType := Real]" } Scale(min := "CV_DATA".HOT_SKID_P03.SCALE_MIN, value := "CV_DATA".HOT_SKID_P03.NORM_OUT, max := "CV_DATA".HOT_SKID_P03.SCALE_MAX, out => "CV_DATA".HOT_SKID_P03.SCALE_OUT)
   END_RUNG
   // the same network as SCL:
   IF 1 THEN
       "CV_DATA".HOT_SKID_P03.NORM_OUT := NORM_X(MIN := "CV_DATA".HOT_SKID_P03.NORM_MIN, VALUE := "CV_DATA".HOT_SKID_P03.OUTPUT_PER, MAX := "CV_DATA".HOT_SKID_P03.NORM_MAX);
       "CV_DATA".HOT_SKID_P03.SCALE_OUT := SCALE_X(MIN := "CV_DATA".HOT_SKID_P03.SCALE_MIN, VALUE := "CV_DATA".HOT_SKID_P03.NORM_OUT, MAX := "CV_DATA".HOT_SKID_P03.SCALE_MAX);
   END_IF;
END_REGION

REGION Network 19: HOT_P03_MANUAL OUTPUT
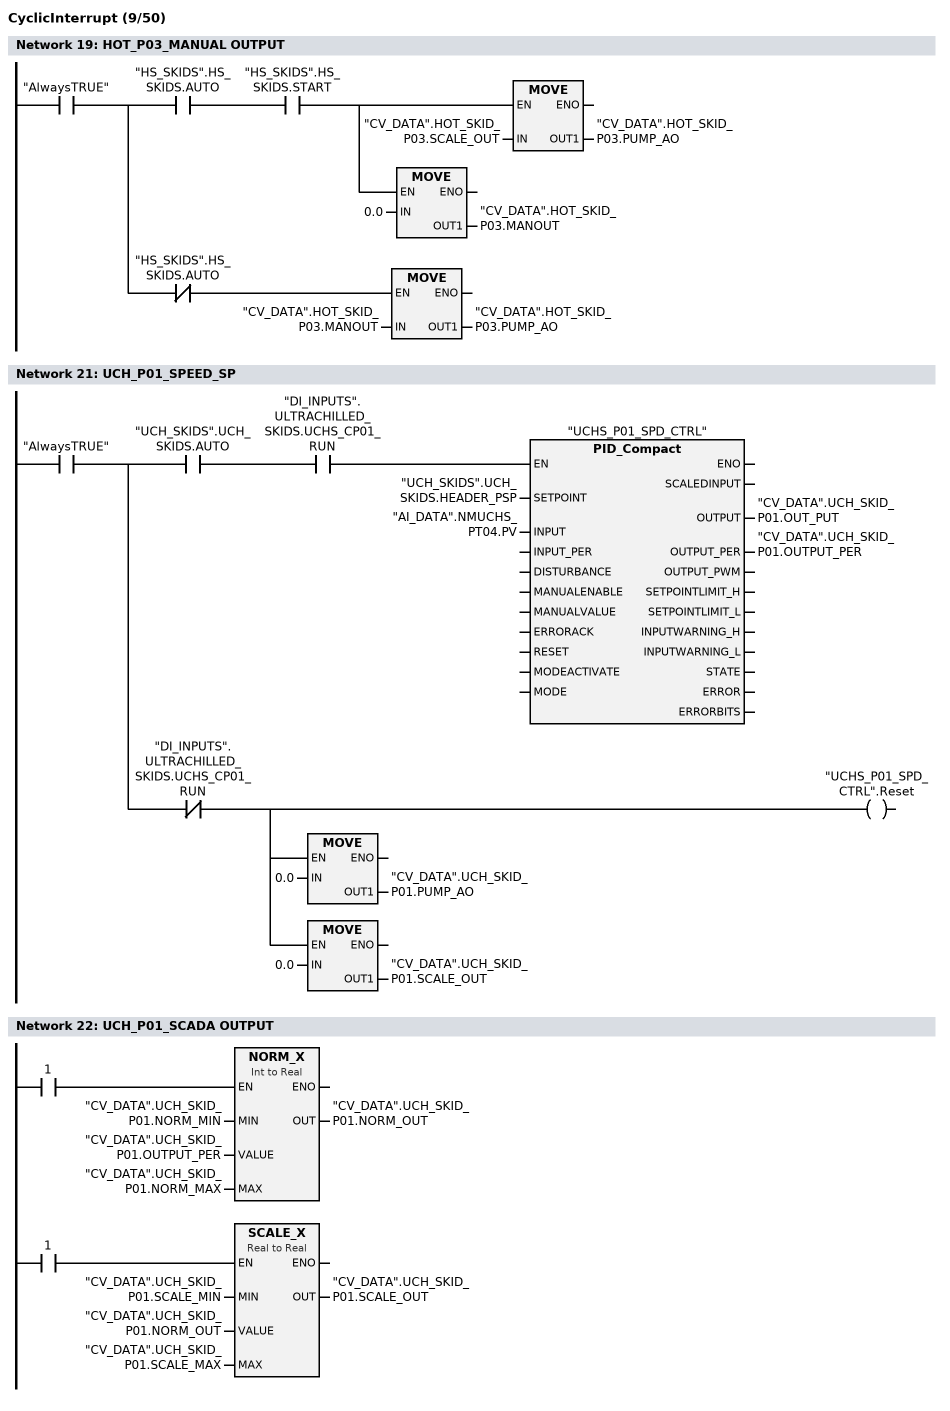
   RUNG wire#powerrail
      Contact( "AlwaysTRUE" )
      wire#w1
      Contact( "HS_SKIDS".HS_SKIDS.AUTO )
      Contact( "HS_SKIDS".HS_SKIDS.START )
      wire#w2
      Move(in := "CV_DATA".HOT_SKID_P03.SCALE_OUT, out1 => "CV_DATA".HOT_SKID_P03.PUMP_AO)
   END_RUNG
   RUNG wire#w2
      Move(in := 0.0, out1 => "CV_DATA".HOT_SKID_P03.MANOUT)
   END_RUNG
   RUNG wire#w1
      I_Contact( "HS_SKIDS".HS_SKIDS.AUTO )
      Move(in := "CV_DATA".HOT_SKID_P03.MANOUT, out1 => "CV_DATA".HOT_SKID_P03.PUMP_AO)
   END_RUNG
   // the same network as SCL:
   IF "AlwaysTRUE" AND "HS_SKIDS".HS_SKIDS.AUTO AND "HS_SKIDS".HS_SKIDS.START THEN
       "CV_DATA".HOT_SKID_P03.PUMP_AO := "CV_DATA".HOT_SKID_P03.SCALE_OUT;
       "CV_DATA".HOT_SKID_P03.MANOUT := 0.0;
   END_IF;
   IF "AlwaysTRUE" AND NOT "HS_SKIDS".HS_SKIDS.AUTO THEN
       "CV_DATA".HOT_SKID_P03.PUMP_AO := "CV_DATA".HOT_SKID_P03.MANOUT;
   END_IF;
END_REGION

REGION Network 21: UCH_P01_SPEED_SP
   RUNG wire#powerrail
      Contact( "AlwaysTRUE" )
      wire#w1
      Contact( "UCH_SKIDS".UCH_SKIDS.AUTO )
      Contact( "DI_INPUTS".ULTRACHILLED_SKIDS.UCHS_CP01_RUN )
      "UCHS_P01_SPD_CTRL".PID_Compact(Setpoint := "UCH_SKIDS".UCH_SKIDS.HEADER_PSP, Input := "AI_DATA".NMUCHS_PT04.PV, Input_PER :=, Disturbance :=, ManualEnable :=, ManualValue :=, ErrorAck :=, Reset :=, ModeActivate :=, Mode :=, ScaledInput =>, Output => "CV_DATA".UCH_SKID_P01.OUT_PUT, Output_PER => "CV_DATA".UCH_SKID_P01.OUTPUT_PER, Output_PWM =>, SetpointLimit_H =>, SetpointLimit_L =>, InputWarning_H =>, InputWarning_L =>, State =>, Error =>, ErrorBits =>)
   END_RUNG
   RUNG wire#w1
      I_Contact( "DI_INPUTS".ULTRACHILLED_SKIDS.UCHS_CP01_RUN )
      wire#w2
      Coil( "UCHS_P01_SPD_CTRL".Reset )
   END_RUNG
   RUNG wire#w2
      Move(in := 0.0, out1 => "CV_DATA".UCH_SKID_P01.PUMP_AO)
   END_RUNG
   RUNG wire#w2
      Move(in := 0.0, out1 => "CV_DATA".UCH_SKID_P01.SCALE_OUT)
   END_RUNG
   // the same network as SCL:
   #_w1 := "AlwaysTRUE";
   IF "AlwaysTRUE" AND "UCH_SKIDS".UCH_SKIDS.AUTO AND "DI_INPUTS".ULTRACHILLED_SKIDS.UCHS_CP01_RUN THEN
       "UCHS_P01_SPD_CTRL"(Setpoint := "UCH_SKIDS".UCH_SKIDS.HEADER_PSP,   // PID_Compact
                           Input := "AI_DATA".NMUCHS_PT04.PV,
                           Output => "CV_DATA".UCH_SKID_P01.OUT_PUT,
                           Output_PER => "CV_DATA".UCH_SKID_P01.OUTPUT_PER);
   END_IF;
   "UCHS_P01_SPD_CTRL".Reset := #_w1 AND NOT "DI_INPUTS".ULTRACHILLED_SKIDS.UCHS_CP01_RUN;
   IF "UCHS_P01_SPD_CTRL".Reset THEN
       "CV_DATA".UCH_SKID_P01.PUMP_AO := 0.0;
       "CV_DATA".UCH_SKID_P01.SCALE_OUT := 0.0;
   END_IF;
END_REGION

REGION Network 22: UCH_P01_SCADA OUTPUT
   RUNG wire#powerrail
      Contact( 1 )
      { S7_Templates := "[SrcType := Int, DestType := Real]" } Normalize(min := "CV_DATA".UCH_SKID_P01.NORM_MIN, value := "CV_DATA".UCH_SKID_P01.OUTPUT_PER, max := "CV_DATA".UCH_SKID_P01.NORM_MAX, out => "CV_DATA".UCH_SKID_P01.NORM_OUT)
   END_RUNG
   RUNG wire#powerrail
      Contact( 1 )
      { S7_Templates := "[SrcType := Real, DestType := Real]" } Scale(min := "CV_DATA".UCH_SKID_P01.SCALE_MIN, value := "CV_DATA".UCH_SKID_P01.NORM_OUT, max := "CV_DATA".UCH_SKID_P01.SCALE_MAX, out => "CV_DATA".UCH_SKID_P01.SCALE_OUT)
   END_RUNG
   // the same network as SCL:
   IF 1 THEN
       "CV_DATA".UCH_SKID_P01.NORM_OUT := NORM_X(MIN := "CV_DATA".UCH_SKID_P01.NORM_MIN, VALUE := "CV_DATA".UCH_SKID_P01.OUTPUT_PER, MAX := "CV_DATA".UCH_SKID_P01.NORM_MAX);
       "CV_DATA".UCH_SKID_P01.SCALE_OUT := SCALE_X(MIN := "CV_DATA".UCH_SKID_P01.SCALE_MIN, VALUE := "CV_DATA".UCH_SKID_P01.NORM_OUT, MAX := "CV_DATA".UCH_SKID_P01.SCALE_MAX);
   END_IF;
END_REGION

REGION Network 23: UCH_P01_MANUAL OUTPUT
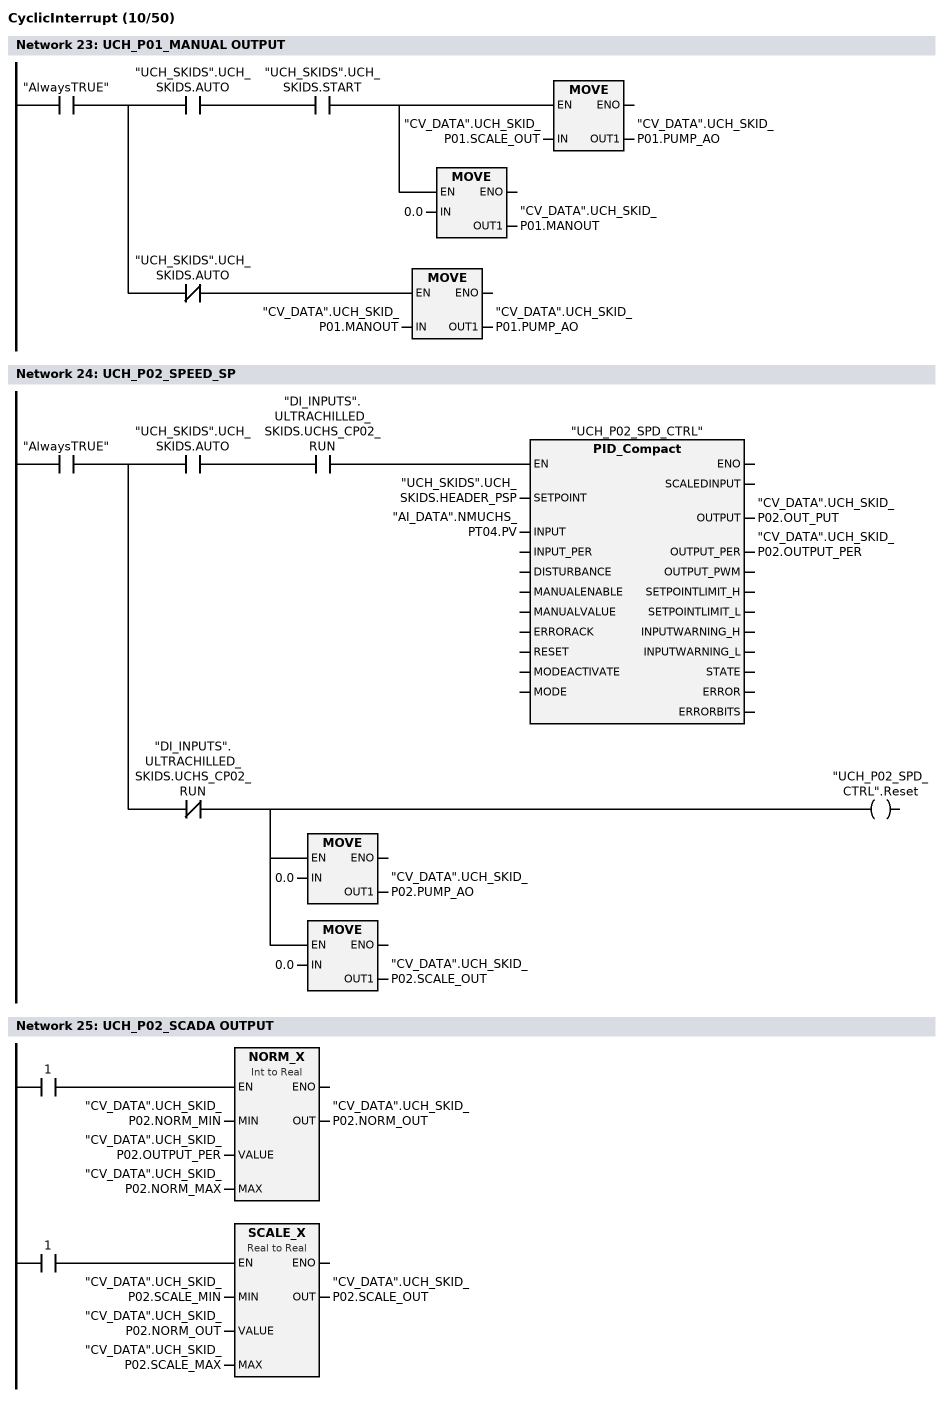
   RUNG wire#powerrail
      Contact( "AlwaysTRUE" )
      wire#w1
      Contact( "UCH_SKIDS".UCH_SKIDS.AUTO )
      Contact( "UCH_SKIDS".UCH_SKIDS.START )
      wire#w2
      Move(in := "CV_DATA".UCH_SKID_P01.SCALE_OUT, out1 => "CV_DATA".UCH_SKID_P01.PUMP_AO)
   END_RUNG
   RUNG wire#w2
      Move(in := 0.0, out1 => "CV_DATA".UCH_SKID_P01.MANOUT)
   END_RUNG
   RUNG wire#w1
      I_Contact( "UCH_SKIDS".UCH_SKIDS.AUTO )
      Move(in := "CV_DATA".UCH_SKID_P01.MANOUT, out1 => "CV_DATA".UCH_SKID_P01.PUMP_AO)
   END_RUNG
   // the same network as SCL:
   IF "AlwaysTRUE" AND "UCH_SKIDS".UCH_SKIDS.AUTO AND "UCH_SKIDS".UCH_SKIDS.START THEN
       "CV_DATA".UCH_SKID_P01.PUMP_AO := "CV_DATA".UCH_SKID_P01.SCALE_OUT;
       "CV_DATA".UCH_SKID_P01.MANOUT := 0.0;
   END_IF;
   IF "AlwaysTRUE" AND NOT "UCH_SKIDS".UCH_SKIDS.AUTO THEN
       "CV_DATA".UCH_SKID_P01.PUMP_AO := "CV_DATA".UCH_SKID_P01.MANOUT;
   END_IF;
END_REGION

REGION Network 24: UCH_P02_SPEED_SP
   RUNG wire#powerrail
      Contact( "AlwaysTRUE" )
      wire#w1
      Contact( "UCH_SKIDS".UCH_SKIDS.AUTO )
      Contact( "DI_INPUTS".ULTRACHILLED_SKIDS.UCHS_CP02_RUN )
      "UCH_P02_SPD_CTRL".PID_Compact(Setpoint := "UCH_SKIDS".UCH_SKIDS.HEADER_PSP, Input := "AI_DATA".NMUCHS_PT04.PV, Input_PER :=, Disturbance :=, ManualEnable :=, ManualValue :=, ErrorAck :=, Reset :=, ModeActivate :=, Mode :=, ScaledInput =>, Output => "CV_DATA".UCH_SKID_P02.OUT_PUT, Output_PER => "CV_DATA".UCH_SKID_P02.OUTPUT_PER, Output_PWM =>, SetpointLimit_H =>, SetpointLimit_L =>, InputWarning_H =>, InputWarning_L =>, State =>, Error =>, ErrorBits =>)
   END_RUNG
   RUNG wire#w1
      I_Contact( "DI_INPUTS".ULTRACHILLED_SKIDS.UCHS_CP02_RUN )
      wire#w2
      Coil( "UCH_P02_SPD_CTRL".Reset )
   END_RUNG
   RUNG wire#w2
      Move(in := 0.0, out1 => "CV_DATA".UCH_SKID_P02.PUMP_AO)
   END_RUNG
   RUNG wire#w2
      Move(in := 0.0, out1 => "CV_DATA".UCH_SKID_P02.SCALE_OUT)
   END_RUNG
   // the same network as SCL:
   #_w1 := "AlwaysTRUE";
   IF "AlwaysTRUE" AND "UCH_SKIDS".UCH_SKIDS.AUTO AND "DI_INPUTS".ULTRACHILLED_SKIDS.UCHS_CP02_RUN THEN
       "UCH_P02_SPD_CTRL"(Setpoint := "UCH_SKIDS".UCH_SKIDS.HEADER_PSP,   // PID_Compact
                          Input := "AI_DATA".NMUCHS_PT04.PV,
                          Output => "CV_DATA".UCH_SKID_P02.OUT_PUT,
                          Output_PER => "CV_DATA".UCH_SKID_P02.OUTPUT_PER);
   END_IF;
   "UCH_P02_SPD_CTRL".Reset := #_w1 AND NOT "DI_INPUTS".ULTRACHILLED_SKIDS.UCHS_CP02_RUN;
   IF "UCH_P02_SPD_CTRL".Reset THEN
       "CV_DATA".UCH_SKID_P02.PUMP_AO := 0.0;
       "CV_DATA".UCH_SKID_P02.SCALE_OUT := 0.0;
   END_IF;
END_REGION

REGION Network 25: UCH_P02_SCADA OUTPUT
   RUNG wire#powerrail
      Contact( 1 )
      { S7_Templates := "[SrcType := Int, DestType := Real]" } Normalize(min := "CV_DATA".UCH_SKID_P02.NORM_MIN, value := "CV_DATA".UCH_SKID_P02.OUTPUT_PER, max := "CV_DATA".UCH_SKID_P02.NORM_MAX, out => "CV_DATA".UCH_SKID_P02.NORM_OUT)
   END_RUNG
   RUNG wire#powerrail
      Contact( 1 )
      { S7_Templates := "[SrcType := Real, DestType := Real]" } Scale(min := "CV_DATA".UCH_SKID_P02.SCALE_MIN, value := "CV_DATA".UCH_SKID_P02.NORM_OUT, max := "CV_DATA".UCH_SKID_P02.SCALE_MAX, out => "CV_DATA".UCH_SKID_P02.SCALE_OUT)
   END_RUNG
   // the same network as SCL:
   IF 1 THEN
       "CV_DATA".UCH_SKID_P02.NORM_OUT := NORM_X(MIN := "CV_DATA".UCH_SKID_P02.NORM_MIN, VALUE := "CV_DATA".UCH_SKID_P02.OUTPUT_PER, MAX := "CV_DATA".UCH_SKID_P02.NORM_MAX);
       "CV_DATA".UCH_SKID_P02.SCALE_OUT := SCALE_X(MIN := "CV_DATA".UCH_SKID_P02.SCALE_MIN, VALUE := "CV_DATA".UCH_SKID_P02.NORM_OUT, MAX := "CV_DATA".UCH_SKID_P02.SCALE_MAX);
   END_IF;
END_REGION

REGION Network 26: UCH_P02_MANUAL OUTPUT
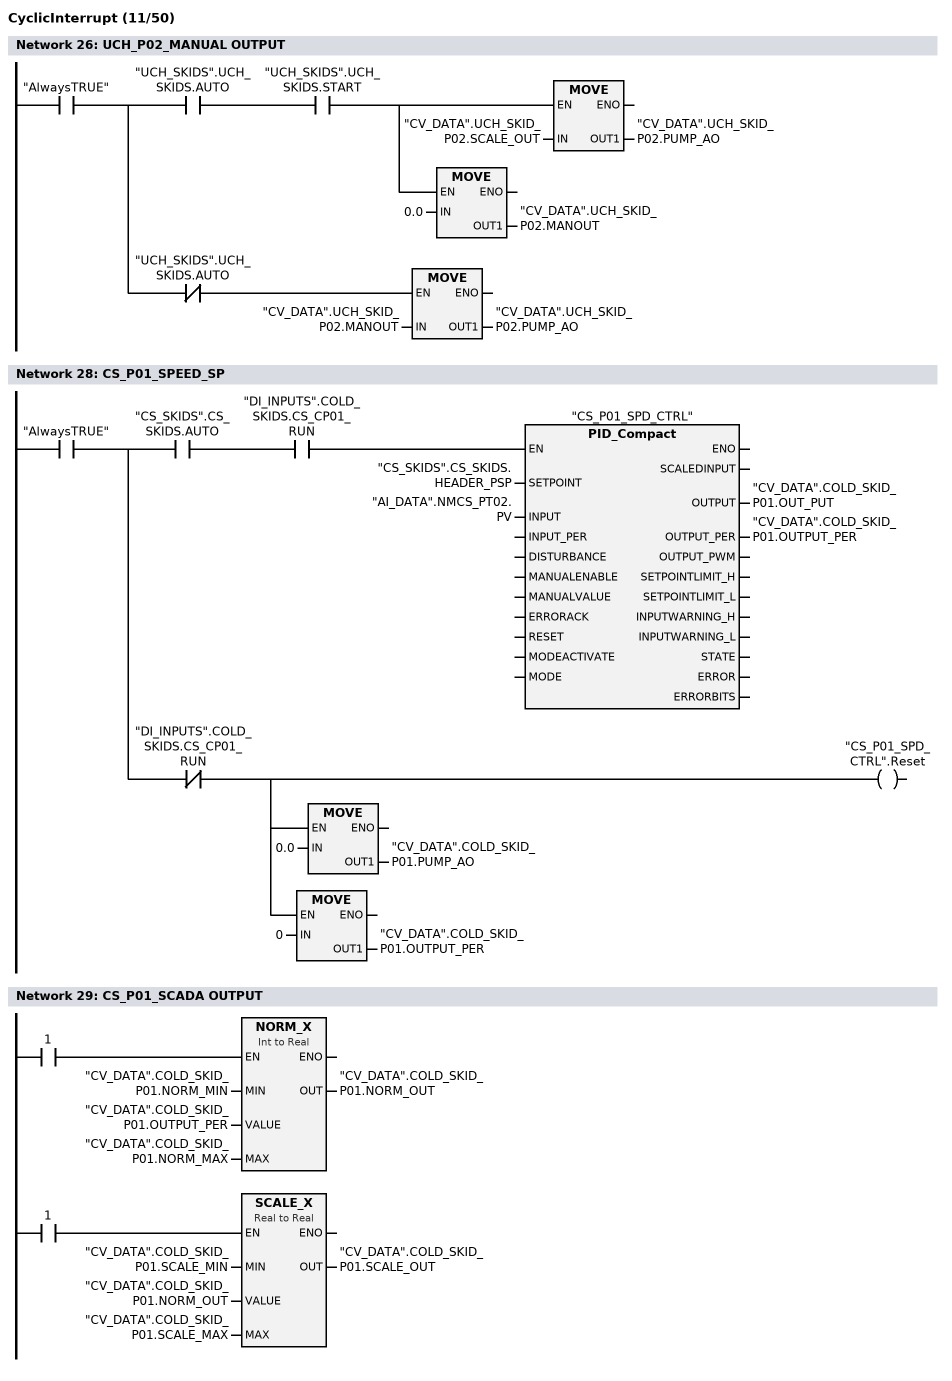
   RUNG wire#powerrail
      Contact( "AlwaysTRUE" )
      wire#w1
      Contact( "UCH_SKIDS".UCH_SKIDS.AUTO )
      Contact( "UCH_SKIDS".UCH_SKIDS.START )
      wire#w2
      Move(in := "CV_DATA".UCH_SKID_P02.SCALE_OUT, out1 => "CV_DATA".UCH_SKID_P02.PUMP_AO)
   END_RUNG
   RUNG wire#w2
      Move(in := 0.0, out1 => "CV_DATA".UCH_SKID_P02.MANOUT)
   END_RUNG
   RUNG wire#w1
      I_Contact( "UCH_SKIDS".UCH_SKIDS.AUTO )
      Move(in := "CV_DATA".UCH_SKID_P02.MANOUT, out1 => "CV_DATA".UCH_SKID_P02.PUMP_AO)
   END_RUNG
   // the same network as SCL:
   IF "AlwaysTRUE" AND "UCH_SKIDS".UCH_SKIDS.AUTO AND "UCH_SKIDS".UCH_SKIDS.START THEN
       "CV_DATA".UCH_SKID_P02.PUMP_AO := "CV_DATA".UCH_SKID_P02.SCALE_OUT;
       "CV_DATA".UCH_SKID_P02.MANOUT := 0.0;
   END_IF;
   IF "AlwaysTRUE" AND NOT "UCH_SKIDS".UCH_SKIDS.AUTO THEN
       "CV_DATA".UCH_SKID_P02.PUMP_AO := "CV_DATA".UCH_SKID_P02.MANOUT;
   END_IF;
END_REGION

REGION Network 28: CS_P01_SPEED_SP
   RUNG wire#powerrail
      Contact( "AlwaysTRUE" )
      wire#w1
      Contact( "CS_SKIDS".CS_SKIDS.AUTO )
      Contact( "DI_INPUTS".COLD_SKIDS.CS_CP01_RUN )
      "CS_P01_SPD_CTRL".PID_Compact(Setpoint := "CS_SKIDS".CS_SKIDS.HEADER_PSP, Input := "AI_DATA".NMCS_PT02.PV, Input_PER :=, Disturbance :=, ManualEnable :=, ManualValue :=, ErrorAck :=, Reset :=, ModeActivate :=, Mode :=, ScaledInput =>, Output => "CV_DATA".COLD_SKID_P01.OUT_PUT, Output_PER => "CV_DATA".COLD_SKID_P01.OUTPUT_PER, Output_PWM =>, SetpointLimit_H =>, SetpointLimit_L =>, InputWarning_H =>, InputWarning_L =>, State =>, Error =>, ErrorBits =>)
   END_RUNG
   RUNG wire#w1
      I_Contact( "DI_INPUTS".COLD_SKIDS.CS_CP01_RUN )
      wire#w2
      Coil( "CS_P01_SPD_CTRL".Reset )
   END_RUNG
   RUNG wire#w2
      Move(in := 0.0, out1 => "CV_DATA".COLD_SKID_P01.PUMP_AO)
   END_RUNG
   RUNG wire#w2
      Move(in := 0, out1 => "CV_DATA".COLD_SKID_P01.OUTPUT_PER)
   END_RUNG
   // the same network as SCL:
   #_w1 := "AlwaysTRUE";
   IF "AlwaysTRUE" AND "CS_SKIDS".CS_SKIDS.AUTO AND "DI_INPUTS".COLD_SKIDS.CS_CP01_RUN THEN
       "CS_P01_SPD_CTRL"(Setpoint := "CS_SKIDS".CS_SKIDS.HEADER_PSP,   // PID_Compact
                         Input := "AI_DATA".NMCS_PT02.PV,
                         Output => "CV_DATA".COLD_SKID_P01.OUT_PUT,
                         Output_PER => "CV_DATA".COLD_SKID_P01.OUTPUT_PER);
   END_IF;
   "CS_P01_SPD_CTRL".Reset := #_w1 AND NOT "DI_INPUTS".COLD_SKIDS.CS_CP01_RUN;
   IF "CS_P01_SPD_CTRL".Reset THEN
       "CV_DATA".COLD_SKID_P01.PUMP_AO := 0.0;
       "CV_DATA".COLD_SKID_P01.OUTPUT_PER := 0;
   END_IF;
END_REGION

REGION Network 29: CS_P01_SCADA OUTPUT
   RUNG wire#powerrail
      Contact( 1 )
      { S7_Templates := "[SrcType := Int, DestType := Real]" } Normalize(min := "CV_DATA".COLD_SKID_P01.NORM_MIN, value := "CV_DATA".COLD_SKID_P01.OUTPUT_PER, max := "CV_DATA".COLD_SKID_P01.NORM_MAX, out => "CV_DATA".COLD_SKID_P01.NORM_OUT)
   END_RUNG
   RUNG wire#powerrail
      Contact( 1 )
      { S7_Templates := "[SrcType := Real, DestType := Real]" } Scale(min := "CV_DATA".COLD_SKID_P01.SCALE_MIN, value := "CV_DATA".COLD_SKID_P01.NORM_OUT, max := "CV_DATA".COLD_SKID_P01.SCALE_MAX, out => "CV_DATA".COLD_SKID_P01.SCALE_OUT)
   END_RUNG
   // the same network as SCL:
   IF 1 THEN
       "CV_DATA".COLD_SKID_P01.NORM_OUT := NORM_X(MIN := "CV_DATA".COLD_SKID_P01.NORM_MIN, VALUE := "CV_DATA".COLD_SKID_P01.OUTPUT_PER, MAX := "CV_DATA".COLD_SKID_P01.NORM_MAX);
       "CV_DATA".COLD_SKID_P01.SCALE_OUT := SCALE_X(MIN := "CV_DATA".COLD_SKID_P01.SCALE_MIN, VALUE := "CV_DATA".COLD_SKID_P01.NORM_OUT, MAX := "CV_DATA".COLD_SKID_P01.SCALE_MAX);
   END_IF;
END_REGION

REGION Network 30: CS_P01_MANUAL OUTPUT
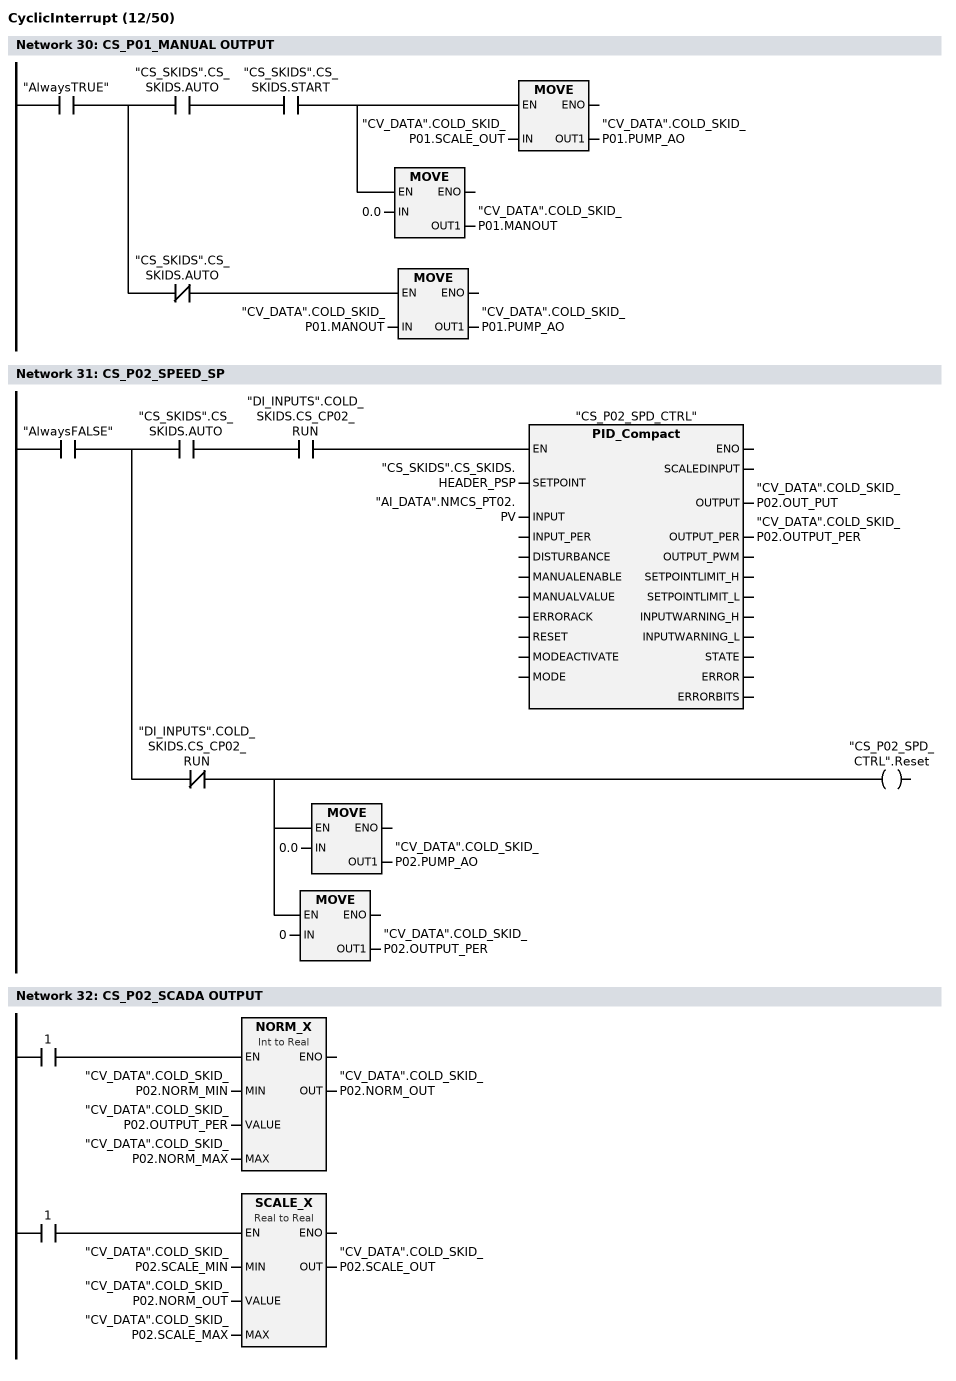
   RUNG wire#powerrail
      Contact( "AlwaysTRUE" )
      wire#w1
      Contact( "CS_SKIDS".CS_SKIDS.AUTO )
      Contact( "CS_SKIDS".CS_SKIDS.START )
      wire#w2
      Move(in := "CV_DATA".COLD_SKID_P01.SCALE_OUT, out1 => "CV_DATA".COLD_SKID_P01.PUMP_AO)
   END_RUNG
   RUNG wire#w2
      Move(in := 0.0, out1 => "CV_DATA".COLD_SKID_P01.MANOUT)
   END_RUNG
   RUNG wire#w1
      I_Contact( "CS_SKIDS".CS_SKIDS.AUTO )
      Move(in := "CV_DATA".COLD_SKID_P01.MANOUT, out1 => "CV_DATA".COLD_SKID_P01.PUMP_AO)
   END_RUNG
   // the same network as SCL:
   IF "AlwaysTRUE" AND "CS_SKIDS".CS_SKIDS.AUTO AND "CS_SKIDS".CS_SKIDS.START THEN
       "CV_DATA".COLD_SKID_P01.PUMP_AO := "CV_DATA".COLD_SKID_P01.SCALE_OUT;
       "CV_DATA".COLD_SKID_P01.MANOUT := 0.0;
   END_IF;
   IF "AlwaysTRUE" AND NOT "CS_SKIDS".CS_SKIDS.AUTO THEN
       "CV_DATA".COLD_SKID_P01.PUMP_AO := "CV_DATA".COLD_SKID_P01.MANOUT;
   END_IF;
END_REGION

REGION Network 31: CS_P02_SPEED_SP
   RUNG wire#powerrail
      Contact( "AlwaysFALSE" )
      wire#w1
      Contact( "CS_SKIDS".CS_SKIDS.AUTO )
      Contact( "DI_INPUTS".COLD_SKIDS.CS_CP02_RUN )
      "CS_P02_SPD_CTRL".PID_Compact(Setpoint := "CS_SKIDS".CS_SKIDS.HEADER_PSP, Input := "AI_DATA".NMCS_PT02.PV, Input_PER :=, Disturbance :=, ManualEnable :=, ManualValue :=, ErrorAck :=, Reset :=, ModeActivate :=, Mode :=, ScaledInput =>, Output => "CV_DATA".COLD_SKID_P02.OUT_PUT, Output_PER => "CV_DATA".COLD_SKID_P02.OUTPUT_PER, Output_PWM =>, SetpointLimit_H =>, SetpointLimit_L =>, InputWarning_H =>, InputWarning_L =>, State =>, Error =>, ErrorBits =>)
   END_RUNG
   RUNG wire#w1
      I_Contact( "DI_INPUTS".COLD_SKIDS.CS_CP02_RUN )
      wire#w2
      Coil( "CS_P02_SPD_CTRL".Reset )
   END_RUNG
   RUNG wire#w2
      Move(in := 0.0, out1 => "CV_DATA".COLD_SKID_P02.PUMP_AO)
   END_RUNG
   RUNG wire#w2
      Move(in := 0, out1 => "CV_DATA".COLD_SKID_P02.OUTPUT_PER)
   END_RUNG
   // the same network as SCL:
   #_w1 := "AlwaysFALSE";
   IF "AlwaysFALSE" AND "CS_SKIDS".CS_SKIDS.AUTO AND "DI_INPUTS".COLD_SKIDS.CS_CP02_RUN THEN
       "CS_P02_SPD_CTRL"(Setpoint := "CS_SKIDS".CS_SKIDS.HEADER_PSP,   // PID_Compact
                         Input := "AI_DATA".NMCS_PT02.PV,
                         Output => "CV_DATA".COLD_SKID_P02.OUT_PUT,
                         Output_PER => "CV_DATA".COLD_SKID_P02.OUTPUT_PER);
   END_IF;
   "CS_P02_SPD_CTRL".Reset := #_w1 AND NOT "DI_INPUTS".COLD_SKIDS.CS_CP02_RUN;
   IF "CS_P02_SPD_CTRL".Reset THEN
       "CV_DATA".COLD_SKID_P02.PUMP_AO := 0.0;
       "CV_DATA".COLD_SKID_P02.OUTPUT_PER := 0;
   END_IF;
END_REGION

REGION Network 32: CS_P02_SCADA OUTPUT
   RUNG wire#powerrail
      Contact( 1 )
      { S7_Templates := "[SrcType := Int, DestType := Real]" } Normalize(min := "CV_DATA".COLD_SKID_P02.NORM_MIN, value := "CV_DATA".COLD_SKID_P02.OUTPUT_PER, max := "CV_DATA".COLD_SKID_P02.NORM_MAX, out => "CV_DATA".COLD_SKID_P02.NORM_OUT)
   END_RUNG
   RUNG wire#powerrail
      Contact( 1 )
      { S7_Templates := "[SrcType := Real, DestType := Real]" } Scale(min := "CV_DATA".COLD_SKID_P02.SCALE_MIN, value := "CV_DATA".COLD_SKID_P02.NORM_OUT, max := "CV_DATA".COLD_SKID_P02.SCALE_MAX, out => "CV_DATA".COLD_SKID_P02.SCALE_OUT)
   END_RUNG
   // the same network as SCL:
   IF 1 THEN
       "CV_DATA".COLD_SKID_P02.NORM_OUT := NORM_X(MIN := "CV_DATA".COLD_SKID_P02.NORM_MIN, VALUE := "CV_DATA".COLD_SKID_P02.OUTPUT_PER, MAX := "CV_DATA".COLD_SKID_P02.NORM_MAX);
       "CV_DATA".COLD_SKID_P02.SCALE_OUT := SCALE_X(MIN := "CV_DATA".COLD_SKID_P02.SCALE_MIN, VALUE := "CV_DATA".COLD_SKID_P02.NORM_OUT, MAX := "CV_DATA".COLD_SKID_P02.SCALE_MAX);
   END_IF;
END_REGION

REGION Network 33: CS_P02_MANUAL OUTPUT
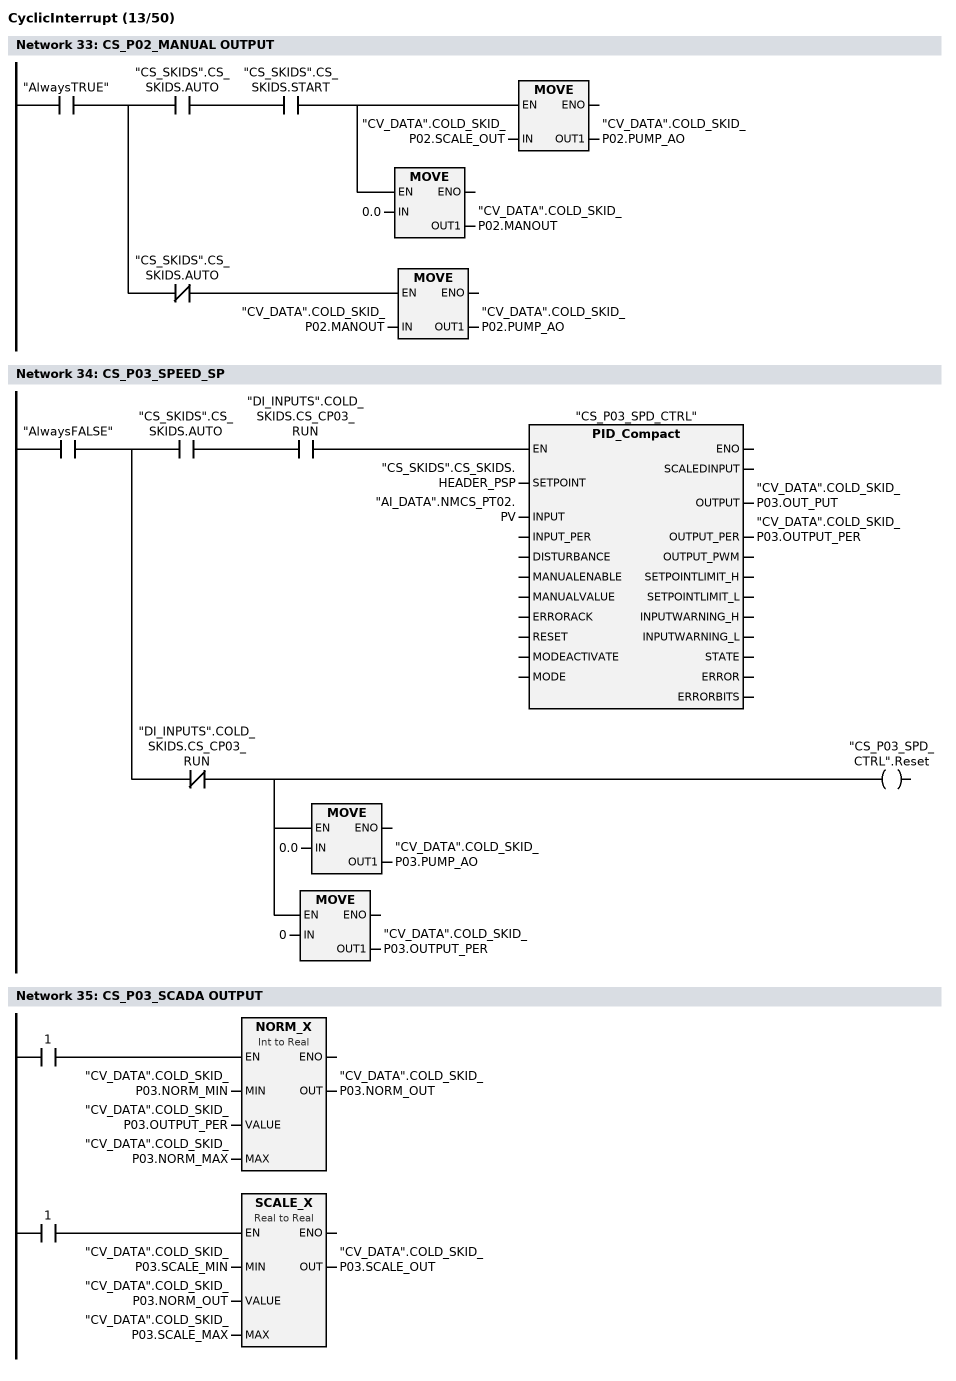
   RUNG wire#powerrail
      Contact( "AlwaysTRUE" )
      wire#w1
      Contact( "CS_SKIDS".CS_SKIDS.AUTO )
      Contact( "CS_SKIDS".CS_SKIDS.START )
      wire#w2
      Move(in := "CV_DATA".COLD_SKID_P02.SCALE_OUT, out1 => "CV_DATA".COLD_SKID_P02.PUMP_AO)
   END_RUNG
   RUNG wire#w2
      Move(in := 0.0, out1 => "CV_DATA".COLD_SKID_P02.MANOUT)
   END_RUNG
   RUNG wire#w1
      I_Contact( "CS_SKIDS".CS_SKIDS.AUTO )
      Move(in := "CV_DATA".COLD_SKID_P02.MANOUT, out1 => "CV_DATA".COLD_SKID_P02.PUMP_AO)
   END_RUNG
   // the same network as SCL:
   IF "AlwaysTRUE" AND "CS_SKIDS".CS_SKIDS.AUTO AND "CS_SKIDS".CS_SKIDS.START THEN
       "CV_DATA".COLD_SKID_P02.PUMP_AO := "CV_DATA".COLD_SKID_P02.SCALE_OUT;
       "CV_DATA".COLD_SKID_P02.MANOUT := 0.0;
   END_IF;
   IF "AlwaysTRUE" AND NOT "CS_SKIDS".CS_SKIDS.AUTO THEN
       "CV_DATA".COLD_SKID_P02.PUMP_AO := "CV_DATA".COLD_SKID_P02.MANOUT;
   END_IF;
END_REGION

REGION Network 34: CS_P03_SPEED_SP
   RUNG wire#powerrail
      Contact( "AlwaysFALSE" )
      wire#w1
      Contact( "CS_SKIDS".CS_SKIDS.AUTO )
      Contact( "DI_INPUTS".COLD_SKIDS.CS_CP03_RUN )
      "CS_P03_SPD_CTRL".PID_Compact(Setpoint := "CS_SKIDS".CS_SKIDS.HEADER_PSP, Input := "AI_DATA".NMCS_PT02.PV, Input_PER :=, Disturbance :=, ManualEnable :=, ManualValue :=, ErrorAck :=, Reset :=, ModeActivate :=, Mode :=, ScaledInput =>, Output => "CV_DATA".COLD_SKID_P03.OUT_PUT, Output_PER => "CV_DATA".COLD_SKID_P03.OUTPUT_PER, Output_PWM =>, SetpointLimit_H =>, SetpointLimit_L =>, InputWarning_H =>, InputWarning_L =>, State =>, Error =>, ErrorBits =>)
   END_RUNG
   RUNG wire#w1
      I_Contact( "DI_INPUTS".COLD_SKIDS.CS_CP03_RUN )
      wire#w2
      Coil( "CS_P03_SPD_CTRL".Reset )
   END_RUNG
   RUNG wire#w2
      Move(in := 0.0, out1 => "CV_DATA".COLD_SKID_P03.PUMP_AO)
   END_RUNG
   RUNG wire#w2
      Move(in := 0, out1 => "CV_DATA".COLD_SKID_P03.OUTPUT_PER)
   END_RUNG
   // the same network as SCL:
   #_w1 := "AlwaysFALSE";
   IF "AlwaysFALSE" AND "CS_SKIDS".CS_SKIDS.AUTO AND "DI_INPUTS".COLD_SKIDS.CS_CP03_RUN THEN
       "CS_P03_SPD_CTRL"(Setpoint := "CS_SKIDS".CS_SKIDS.HEADER_PSP,   // PID_Compact
                         Input := "AI_DATA".NMCS_PT02.PV,
                         Output => "CV_DATA".COLD_SKID_P03.OUT_PUT,
                         Output_PER => "CV_DATA".COLD_SKID_P03.OUTPUT_PER);
   END_IF;
   "CS_P03_SPD_CTRL".Reset := #_w1 AND NOT "DI_INPUTS".COLD_SKIDS.CS_CP03_RUN;
   IF "CS_P03_SPD_CTRL".Reset THEN
       "CV_DATA".COLD_SKID_P03.PUMP_AO := 0.0;
       "CV_DATA".COLD_SKID_P03.OUTPUT_PER := 0;
   END_IF;
END_REGION

REGION Network 35: CS_P03_SCADA OUTPUT
   RUNG wire#powerrail
      Contact( 1 )
      { S7_Templates := "[SrcType := Int, DestType := Real]" } Normalize(min := "CV_DATA".COLD_SKID_P03.NORM_MIN, value := "CV_DATA".COLD_SKID_P03.OUTPUT_PER, max := "CV_DATA".COLD_SKID_P03.NORM_MAX, out => "CV_DATA".COLD_SKID_P03.NORM_OUT)
   END_RUNG
   RUNG wire#powerrail
      Contact( 1 )
      { S7_Templates := "[SrcType := Real, DestType := Real]" } Scale(min := "CV_DATA".COLD_SKID_P03.SCALE_MIN, value := "CV_DATA".COLD_SKID_P03.NORM_OUT, max := "CV_DATA".COLD_SKID_P03.SCALE_MAX, out => "CV_DATA".COLD_SKID_P03.SCALE_OUT)
   END_RUNG
   // the same network as SCL:
   IF 1 THEN
       "CV_DATA".COLD_SKID_P03.NORM_OUT := NORM_X(MIN := "CV_DATA".COLD_SKID_P03.NORM_MIN, VALUE := "CV_DATA".COLD_SKID_P03.OUTPUT_PER, MAX := "CV_DATA".COLD_SKID_P03.NORM_MAX);
       "CV_DATA".COLD_SKID_P03.SCALE_OUT := SCALE_X(MIN := "CV_DATA".COLD_SKID_P03.SCALE_MIN, VALUE := "CV_DATA".COLD_SKID_P03.NORM_OUT, MAX := "CV_DATA".COLD_SKID_P03.SCALE_MAX);
   END_IF;
END_REGION

REGION Network 36: CS_P03_MANUAL OUTPUT
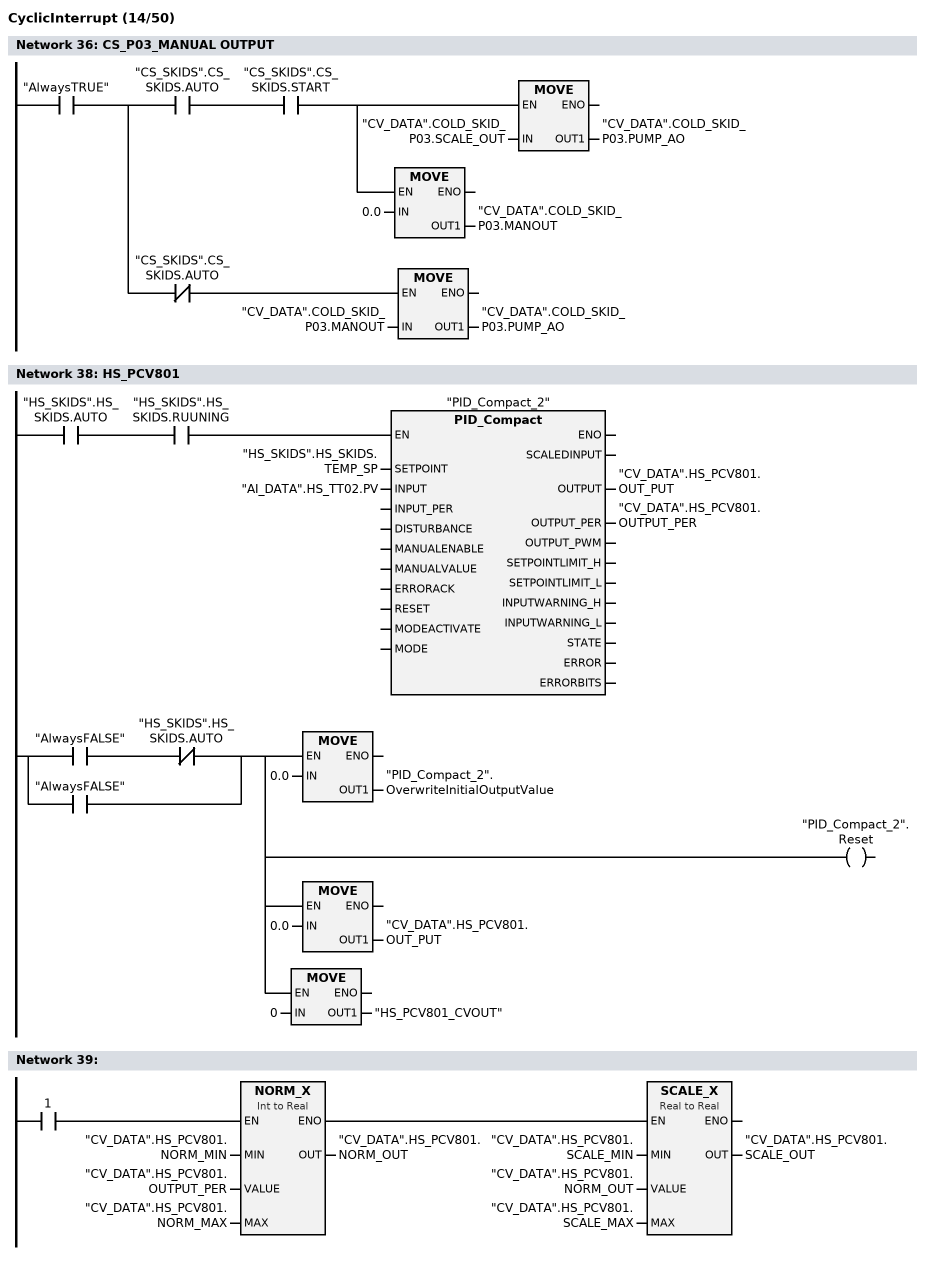
   RUNG wire#powerrail
      Contact( "AlwaysTRUE" )
      wire#w1
      Contact( "CS_SKIDS".CS_SKIDS.AUTO )
      Contact( "CS_SKIDS".CS_SKIDS.START )
      wire#w2
      Move(in := "CV_DATA".COLD_SKID_P03.SCALE_OUT, out1 => "CV_DATA".COLD_SKID_P03.PUMP_AO)
   END_RUNG
   RUNG wire#w2
      Move(in := 0.0, out1 => "CV_DATA".COLD_SKID_P03.MANOUT)
   END_RUNG
   RUNG wire#w1
      I_Contact( "CS_SKIDS".CS_SKIDS.AUTO )
      Move(in := "CV_DATA".COLD_SKID_P03.MANOUT, out1 => "CV_DATA".COLD_SKID_P03.PUMP_AO)
   END_RUNG
   // the same network as SCL:
   IF "AlwaysTRUE" AND "CS_SKIDS".CS_SKIDS.AUTO AND "CS_SKIDS".CS_SKIDS.START THEN
       "CV_DATA".COLD_SKID_P03.PUMP_AO := "CV_DATA".COLD_SKID_P03.SCALE_OUT;
       "CV_DATA".COLD_SKID_P03.MANOUT := 0.0;
   END_IF;
   IF "AlwaysTRUE" AND NOT "CS_SKIDS".CS_SKIDS.AUTO THEN
       "CV_DATA".COLD_SKID_P03.PUMP_AO := "CV_DATA".COLD_SKID_P03.MANOUT;
   END_IF;
END_REGION

REGION Network 38: HS_PCV801
   RUNG wire#powerrail
      Contact( "HS_SKIDS".HS_SKIDS.AUTO )
      Contact( "HS_SKIDS".HS_SKIDS.RUUNING )
      "PID_Compact_2".PID_Compact(Setpoint := "HS_SKIDS".HS_SKIDS.TEMP_SP, Input := "AI_DATA".HS_TT02.PV, Input_PER :=, Disturbance :=, ManualEnable :=, ManualValue :=, ErrorAck :=, Reset :=, ModeActivate :=, Mode :=, ScaledInput =>, Output => "CV_DATA".HS_PCV801.OUT_PUT, Output_PER => "CV_DATA".HS_PCV801.OUTPUT_PER, Output_PWM =>, SetpointLimit_H =>, SetpointLimit_L =>, InputWarning_H =>, InputWarning_L =>, State =>, Error =>, ErrorBits =>)
   END_RUNG
   RUNG wire#powerrail
      Contact( "AlwaysFALSE" )
      I_Contact( "HS_SKIDS".HS_SKIDS.AUTO )
      wire#w1
      Move(in := 0.0, out1 => "PID_Compact_2".OverwriteInitialOutputValue)
   END_RUNG
   RUNG wire#powerrail
      Contact( "AlwaysFALSE" )
   END_RUNG wire#w1
   RUNG wire#w1
      Coil( "PID_Compact_2".Reset )
   END_RUNG
   RUNG wire#w1
      Move(in := 0.0, out1 => "CV_DATA".HS_PCV801.OUT_PUT)
   END_RUNG
   RUNG wire#w1
      Move(in := 0, out1 => "HS_PCV801_CVOUT")
   END_RUNG
   // the same network as SCL:
   IF "HS_SKIDS".HS_SKIDS.AUTO AND "HS_SKIDS".HS_SKIDS.RUUNING THEN
       "PID_Compact_2"(Setpoint := "HS_SKIDS".HS_SKIDS.TEMP_SP,   // PID_Compact
                       Input := "AI_DATA".HS_TT02.PV,
                       Output => "CV_DATA".HS_PCV801.OUT_PUT,
                       Output_PER => "CV_DATA".HS_PCV801.OUTPUT_PER);
   END_IF;
   #_w1 := ("AlwaysFALSE" AND NOT "HS_SKIDS".HS_SKIDS.AUTO) OR "AlwaysFALSE";
   IF #_w1 THEN "PID_Compact_2".OverwriteInitialOutputValue := 0.0; END_IF;
   "PID_Compact_2".Reset := #_w1;
   IF #_w1 THEN
       "CV_DATA".HS_PCV801.OUT_PUT := 0.0;
       "HS_PCV801_CVOUT" := 0;
   END_IF;
END_REGION

REGION Network 39
   RUNG wire#powerrail
      Contact( 1 )
      { S7_Templates := "[SrcType := Int, DestType := Real]" } Normalize(min := "CV_DATA".HS_PCV801.NORM_MIN, value := "CV_DATA".HS_PCV801.OUTPUT_PER, max := "CV_DATA".HS_PCV801.NORM_MAX, out => "CV_DATA".HS_PCV801.NORM_OUT)
      { S7_Templates := "[SrcType := Real, DestType := Real]" } Scale(min := "CV_DATA".HS_PCV801.SCALE_MIN, value := "CV_DATA".HS_PCV801.NORM_OUT, max := "CV_DATA".HS_PCV801.SCALE_MAX, out => "CV_DATA".HS_PCV801.SCALE_OUT)
   END_RUNG
   // the same network as SCL:
   IF 1 THEN
       "CV_DATA".HS_PCV801.NORM_OUT := NORM_X(MIN := "CV_DATA".HS_PCV801.NORM_MIN, VALUE := "CV_DATA".HS_PCV801.OUTPUT_PER, MAX := "CV_DATA".HS_PCV801.NORM_MAX);
       "CV_DATA".HS_PCV801.SCALE_OUT := SCALE_X(MIN := "CV_DATA".HS_PCV801.SCALE_MIN, VALUE := "CV_DATA".HS_PCV801.NORM_OUT, MAX := "CV_DATA".HS_PCV801.SCALE_MAX);
   END_IF;
END_REGION

REGION Network 40
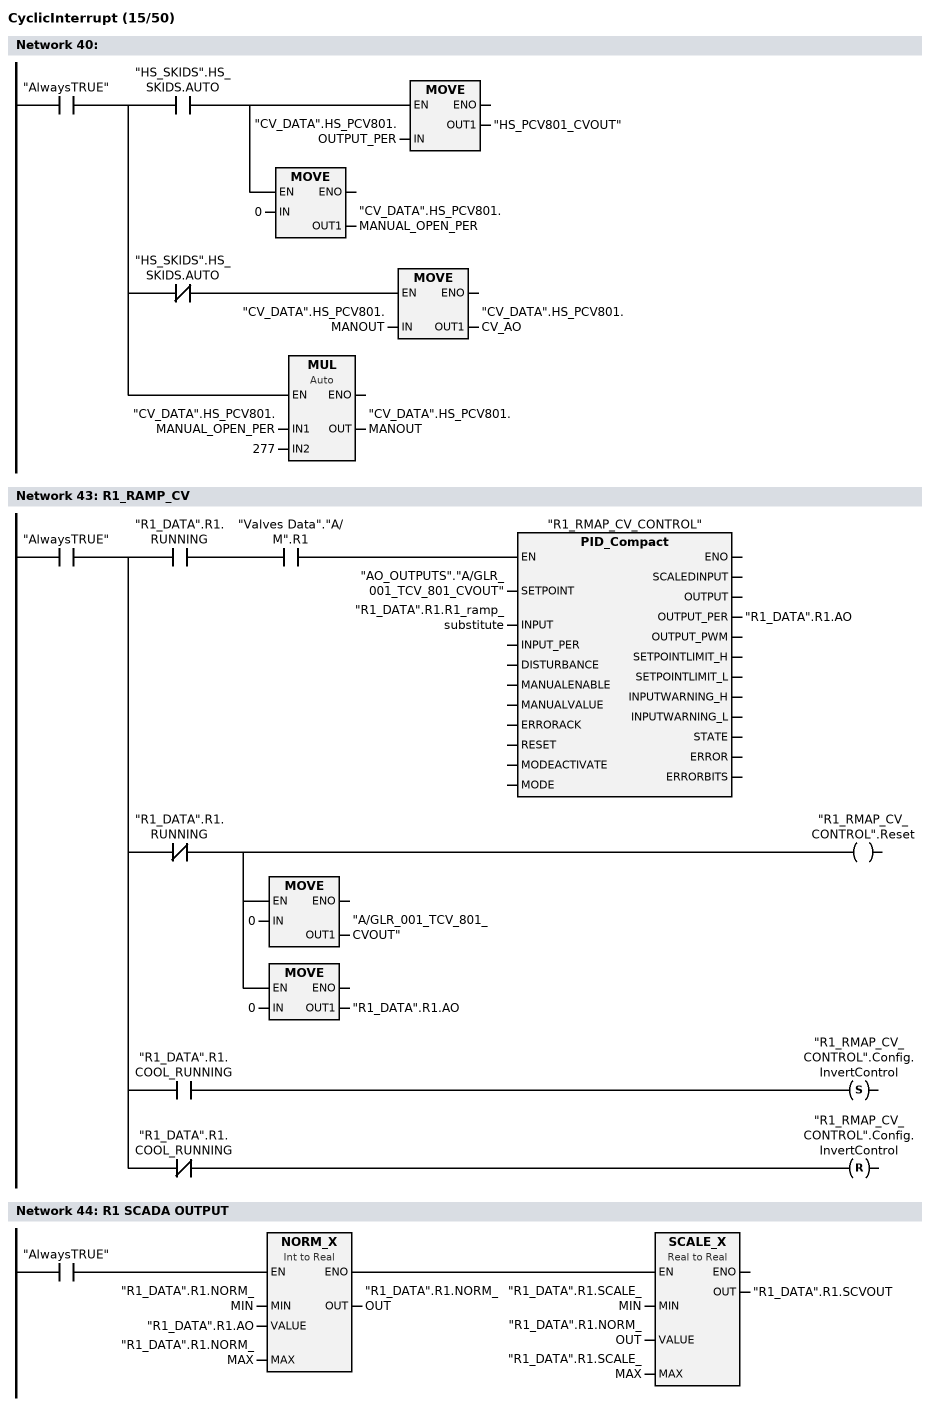
   RUNG wire#powerrail
      Contact( "AlwaysTRUE" )
      wire#w1
      Contact( "HS_SKIDS".HS_SKIDS.AUTO )
      wire#w2
      Move(in := "CV_DATA".HS_PCV801.OUTPUT_PER, out1 => "HS_PCV801_CVOUT")
   END_RUNG
   RUNG wire#w2
      Move(in := 0, out1 => "CV_DATA".HS_PCV801.MANUAL_OPEN_PER)
   END_RUNG
   RUNG wire#w1
      I_Contact( "HS_SKIDS".HS_SKIDS.AUTO )
      Move(in := "CV_DATA".HS_PCV801.MANOUT, out1 => "CV_DATA".HS_PCV801.CV_AO)
   END_RUNG
   RUNG wire#w1
      Mul(in1 := "CV_DATA".HS_PCV801.MANUAL_OPEN_PER, in2 := 277, out => "CV_DATA".HS_PCV801.MANOUT)
   END_RUNG
   // the same network as SCL:
   IF "AlwaysTRUE" AND "HS_SKIDS".HS_SKIDS.AUTO THEN
       "HS_PCV801_CVOUT" := "CV_DATA".HS_PCV801.OUTPUT_PER;
       "CV_DATA".HS_PCV801.MANUAL_OPEN_PER := 0;
   END_IF;
   IF "AlwaysTRUE" AND NOT "HS_SKIDS".HS_SKIDS.AUTO THEN
       "CV_DATA".HS_PCV801.CV_AO := "CV_DATA".HS_PCV801.MANOUT;
   END_IF;
   IF "AlwaysTRUE" THEN "CV_DATA".HS_PCV801.MANOUT := "CV_DATA".HS_PCV801.MANUAL_OPEN_PER * 277; END_IF;
END_REGION

REGION Network 43: R1_RAMP_CV
   RUNG wire#powerrail
      Contact( "AlwaysTRUE" )
      wire#w1
      Contact( "R1_DATA".R1.RUNNING )
      Contact( "Valves Data"."A/M".R1 )
      "R1_RMAP_CV_CONTROL".PID_Compact(Setpoint := "AO_OUTPUTS"."A/GLR_001_TCV_801_CVOUT", Input := "R1_DATA".R1.R1_ramp_substitute, Input_PER :=, Disturbance :=, ManualEnable :=, ManualValue :=, ErrorAck :=, Reset :=, ModeActivate :=, Mode :=, ScaledInput =>, Output =>, Output_PER => "R1_DATA".R1.AO, Output_PWM =>, SetpointLimit_H =>, SetpointLimit_L =>, InputWarning_H =>, InputWarning_L =>, State =>, Error =>, ErrorBits =>)
   END_RUNG
   RUNG wire#w1
      I_Contact( "R1_DATA".R1.RUNNING )
      wire#w2
      Coil( "R1_RMAP_CV_CONTROL".Reset )
   END_RUNG
   RUNG wire#w2
      Move(in := 0, out1 => "A/GLR_001_TCV_801_CVOUT")
   END_RUNG
   RUNG wire#w2
      Move(in := 0, out1 => "R1_DATA".R1.AO)
   END_RUNG
   RUNG wire#w1
      Contact( "R1_DATA".R1.COOL_RUNNING )
      S_Coil( "R1_RMAP_CV_CONTROL".Config.InvertControl )
   END_RUNG
   RUNG wire#w1
      I_Contact( "R1_DATA".R1.COOL_RUNNING )
      R_Coil( "R1_RMAP_CV_CONTROL".Config.InvertControl )
   END_RUNG
   // the same network as SCL:
   #_w1 := "AlwaysTRUE";
   IF "AlwaysTRUE" AND "R1_DATA".R1.RUNNING AND "Valves Data"."A/M".R1 THEN
       "R1_RMAP_CV_CONTROL"(Setpoint := "AO_OUTPUTS"."A/GLR_001_TCV_801_CVOUT",   // PID_Compact
                            Input := "R1_DATA".R1.R1_ramp_substitute,
                            Output_PER => "R1_DATA".R1.AO);
   END_IF;
   "R1_RMAP_CV_CONTROL".Reset := #_w1 AND NOT "R1_DATA".R1.RUNNING;
   IF "R1_RMAP_CV_CONTROL".Reset THEN
       "A/GLR_001_TCV_801_CVOUT" := 0;
       "R1_DATA".R1.AO := 0;
   END_IF;
   IF #_w1 AND "R1_DATA".R1.COOL_RUNNING THEN "R1_RMAP_CV_CONTROL".Config.InvertControl := TRUE; END_IF;
   IF #_w1 AND NOT "R1_DATA".R1.COOL_RUNNING THEN "R1_RMAP_CV_CONTROL".Config.InvertControl := FALSE; END_IF;
END_REGION

REGION Network 44: R1 SCADA OUTPUT
   RUNG wire#powerrail
      Contact( "AlwaysTRUE" )
      { S7_Templates := "[SrcType := Int, DestType := Real]" } Normalize(min := "R1_DATA".R1.NORM_MIN, value := "R1_DATA".R1.AO, max := "R1_DATA".R1.NORM_MAX, out => "R1_DATA".R1.NORM_OUT)
      { S7_Templates := "[SrcType := Real, DestType := Real]" } Scale(min := "R1_DATA".R1.SCALE_MIN, value := "R1_DATA".R1.NORM_OUT, max := "R1_DATA".R1.SCALE_MAX, out => "R1_DATA".R1.SCVOUT)
   END_RUNG
   // the same network as SCL:
   IF "AlwaysTRUE" THEN
       "R1_DATA".R1.NORM_OUT := NORM_X(MIN := "R1_DATA".R1.NORM_MIN, VALUE := "R1_DATA".R1.AO, MAX := "R1_DATA".R1.NORM_MAX);
       "R1_DATA".R1.SCVOUT := SCALE_X(MIN := "R1_DATA".R1.SCALE_MIN, VALUE := "R1_DATA".R1.NORM_OUT, MAX := "R1_DATA".R1.SCALE_MAX);
   END_IF;
END_REGION

REGION Network 45: R1 AUTO/MANUAL OUTPUT
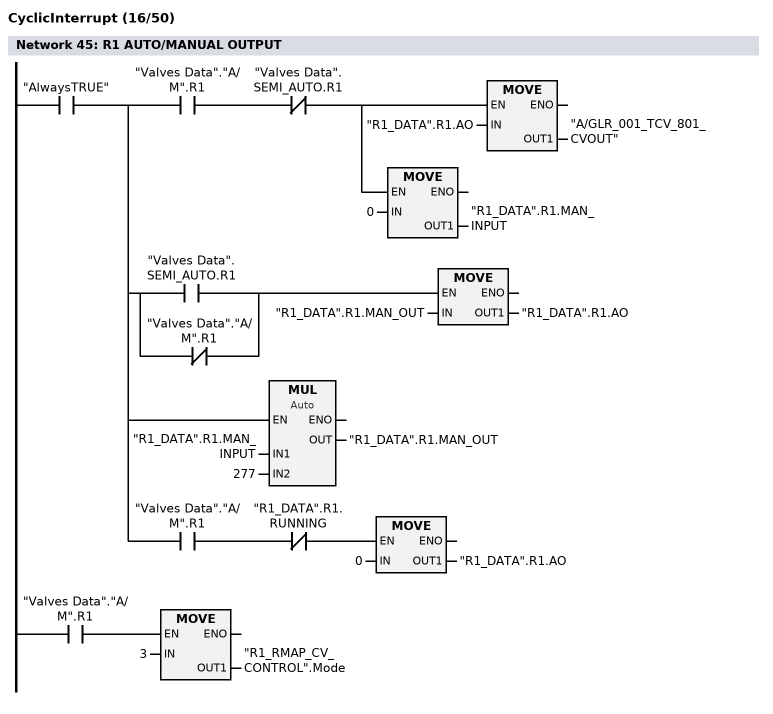
   RUNG wire#powerrail
      Contact( "AlwaysTRUE" )
      wire#w1
      Contact( "Valves Data"."A/M".R1 )
      I_Contact( "Valves Data".SEMI_AUTO.R1 )
      wire#w2
      Move(in := "R1_DATA".R1.AO, out1 => "A/GLR_001_TCV_801_CVOUT")
   END_RUNG
   RUNG wire#w2
      Move(in := 0, out1 => "R1_DATA".R1.MAN_INPUT)
   END_RUNG
   RUNG wire#w1
      Contact( "Valves Data".SEMI_AUTO.R1 )
      wire#w3
      Move(in := "R1_DATA".R1.MAN_OUT, out1 => "R1_DATA".R1.AO)
   END_RUNG
   RUNG wire#w1
      I_Contact( "Valves Data"."A/M".R1 )
   END_RUNG wire#w3
   RUNG wire#w1
      Mul(in1 := "R1_DATA".R1.MAN_INPUT, in2 := 277, out => "R1_DATA".R1.MAN_OUT)
   END_RUNG
   RUNG wire#w1
      Contact( "Valves Data"."A/M".R1 )
      I_Contact( "R1_DATA".R1.RUNNING )
      Move(in := 0, out1 => "R1_DATA".R1.AO)
   END_RUNG
   RUNG wire#powerrail
      Contact( "Valves Data"."A/M".R1 )
      Move(in := 3, out1 => "R1_RMAP_CV_CONTROL".Mode)
   END_RUNG
   // the same network as SCL:
   IF "AlwaysTRUE" AND "Valves Data"."A/M".R1 AND NOT "Valves Data".SEMI_AUTO.R1 THEN
       "A/GLR_001_TCV_801_CVOUT" := "R1_DATA".R1.AO;
       "R1_DATA".R1.MAN_INPUT := 0;
   END_IF;
   IF "AlwaysTRUE" AND ("Valves Data".SEMI_AUTO.R1 OR NOT "Valves Data"."A/M".R1) THEN
       "R1_DATA".R1.AO := "R1_DATA".R1.MAN_OUT;
   END_IF;
   IF "AlwaysTRUE" THEN "R1_DATA".R1.MAN_OUT := "R1_DATA".R1.MAN_INPUT * 277; END_IF;
   IF "AlwaysTRUE" AND "Valves Data"."A/M".R1 AND NOT "R1_DATA".R1.RUNNING THEN "R1_DATA".R1.AO := 0; END_IF;
   IF "Valves Data"."A/M".R1 THEN "R1_RMAP_CV_CONTROL".Mode := 3; END_IF;
END_REGION

REGION Network 46: R2_RAMP_CV
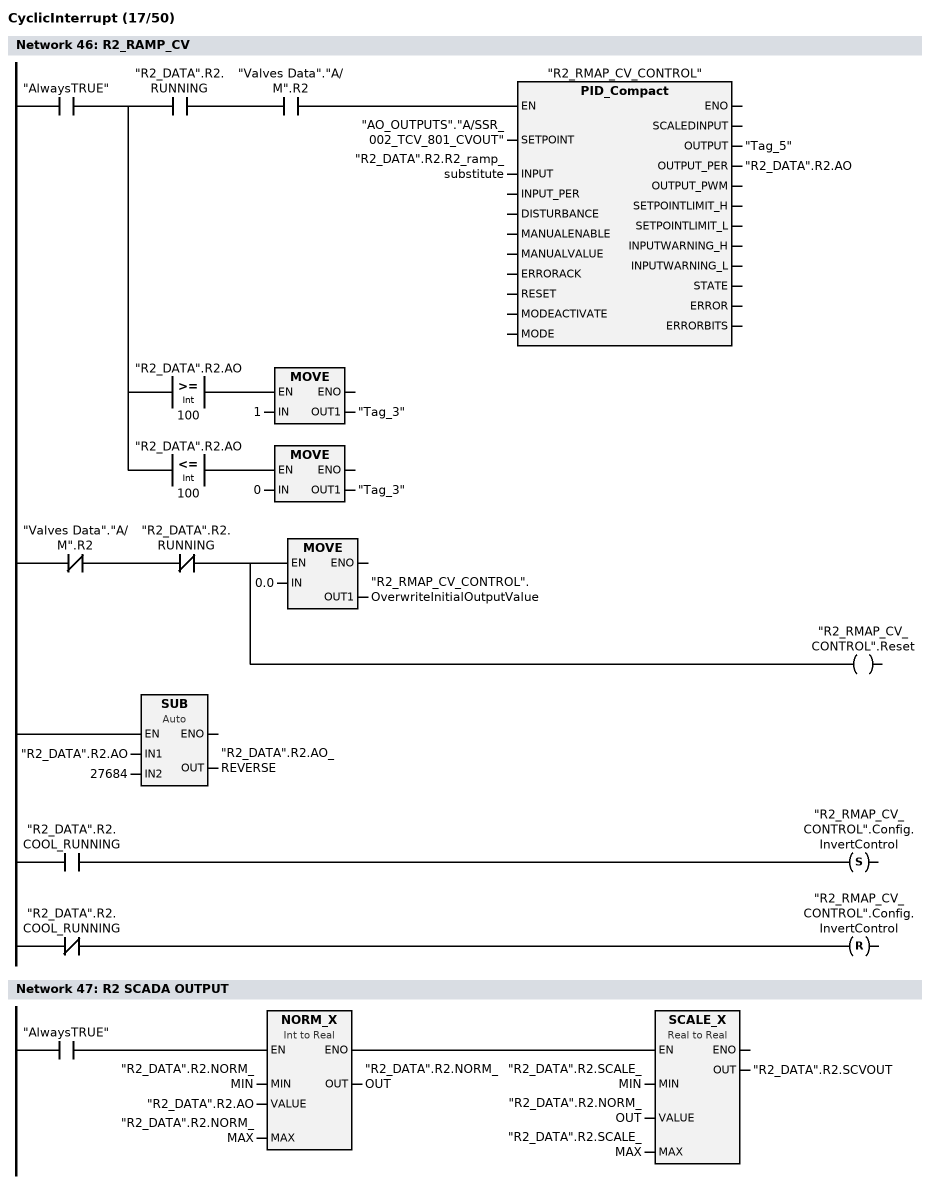
   RUNG wire#powerrail
      Contact( "AlwaysTRUE" )
      wire#w1
      Contact( "R2_DATA".R2.RUNNING )
      Contact( "Valves Data"."A/M".R2 )
      "R2_RMAP_CV_CONTROL".PID_Compact(Setpoint := "AO_OUTPUTS"."A/SSR_002_TCV_801_CVOUT", Input := "R2_DATA".R2.R2_ramp_substitute, Input_PER :=, Disturbance :=, ManualEnable :=, ManualValue :=, ErrorAck :=, Reset :=, ModeActivate :=, Mode :=, ScaledInput =>, Output => "Tag_5", Output_PER => "R2_DATA".R2.AO, Output_PWM =>, SetpointLimit_H =>, SetpointLimit_L =>, InputWarning_H =>, InputWarning_L =>, State =>, Error =>, ErrorBits =>)
   END_RUNG
   RUNG wire#w1
      { S7_Templates := "SrcType := Int" } GE_Contact(in1 := "R2_DATA".R2.AO, in2 := 100)
      Move(in := 1, out1 => "Tag_3")
   END_RUNG
   RUNG wire#w1
      { S7_Templates := "SrcType := Int" } LE_Contact(in1 := "R2_DATA".R2.AO, in2 := 100)
      Move(in := 0, out1 => "Tag_3")
   END_RUNG
   RUNG wire#powerrail
      I_Contact( "Valves Data"."A/M".R2 )
      I_Contact( "R2_DATA".R2.RUNNING )
      wire#w2
      Move(in := 0.0, out1 => "R2_RMAP_CV_CONTROL".OverwriteInitialOutputValue)
   END_RUNG
   RUNG wire#w2
      Coil( "R2_RMAP_CV_CONTROL".Reset )
   END_RUNG
   RUNG wire#powerrail
      Sub(in1 := "R2_DATA".R2.AO, in2 := 27684, out => "R2_DATA".R2.AO_REVERSE)
   END_RUNG
   RUNG wire#powerrail
      Contact( "R2_DATA".R2.COOL_RUNNING )
      S_Coil( "R2_RMAP_CV_CONTROL".Config.InvertControl )
   END_RUNG
   RUNG wire#powerrail
      I_Contact( "R2_DATA".R2.COOL_RUNNING )
      R_Coil( "R2_RMAP_CV_CONTROL".Config.InvertControl )
   END_RUNG
   // the same network as SCL:
   #_w1 := "AlwaysTRUE";
   IF "AlwaysTRUE" AND "R2_DATA".R2.RUNNING AND "Valves Data"."A/M".R2 THEN
       "R2_RMAP_CV_CONTROL"(Setpoint := "AO_OUTPUTS"."A/SSR_002_TCV_801_CVOUT",   // PID_Compact
                            Input := "R2_DATA".R2.R2_ramp_substitute,
                            Output => "Tag_5",
                            Output_PER => "R2_DATA".R2.AO);
   END_IF;
   IF #_w1 AND ("R2_DATA".R2.AO >= 100) THEN "Tag_3" := 1; END_IF;
   IF #_w1 AND ("R2_DATA".R2.AO <= 100) THEN "Tag_3" := 0; END_IF;
   #_w2 := NOT "Valves Data"."A/M".R2 AND NOT "R2_DATA".R2.RUNNING;
   IF #_w2 THEN "R2_RMAP_CV_CONTROL".OverwriteInitialOutputValue := 0.0; END_IF;
   "R2_RMAP_CV_CONTROL".Reset := #_w2;
   "R2_DATA".R2.AO_REVERSE := "R2_DATA".R2.AO - 27684;
   IF "R2_DATA".R2.COOL_RUNNING THEN "R2_RMAP_CV_CONTROL".Config.InvertControl := TRUE; END_IF;
   IF NOT "R2_DATA".R2.COOL_RUNNING THEN "R2_RMAP_CV_CONTROL".Config.InvertControl := FALSE; END_IF;
END_REGION

REGION Network 47: R2 SCADA OUTPUT
   RUNG wire#powerrail
      Contact( "AlwaysTRUE" )
      { S7_Templates := "[SrcType := Int, DestType := Real]" } Normalize(min := "R2_DATA".R2.NORM_MIN, value := "R2_DATA".R2.AO, max := "R2_DATA".R2.NORM_MAX, out => "R2_DATA".R2.NORM_OUT)
      { S7_Templates := "[SrcType := Real, DestType := Real]" } Scale(min := "R2_DATA".R2.SCALE_MIN, value := "R2_DATA".R2.NORM_OUT, max := "R2_DATA".R2.SCALE_MAX, out => "R2_DATA".R2.SCVOUT)
   END_RUNG
   // the same network as SCL:
   IF "AlwaysTRUE" THEN
       "R2_DATA".R2.NORM_OUT := NORM_X(MIN := "R2_DATA".R2.NORM_MIN, VALUE := "R2_DATA".R2.AO, MAX := "R2_DATA".R2.NORM_MAX);
       "R2_DATA".R2.SCVOUT := SCALE_X(MIN := "R2_DATA".R2.SCALE_MIN, VALUE := "R2_DATA".R2.NORM_OUT, MAX := "R2_DATA".R2.SCALE_MAX);
   END_IF;
END_REGION

REGION Network 48: R2 AUTO/MANUAL OUTPUT
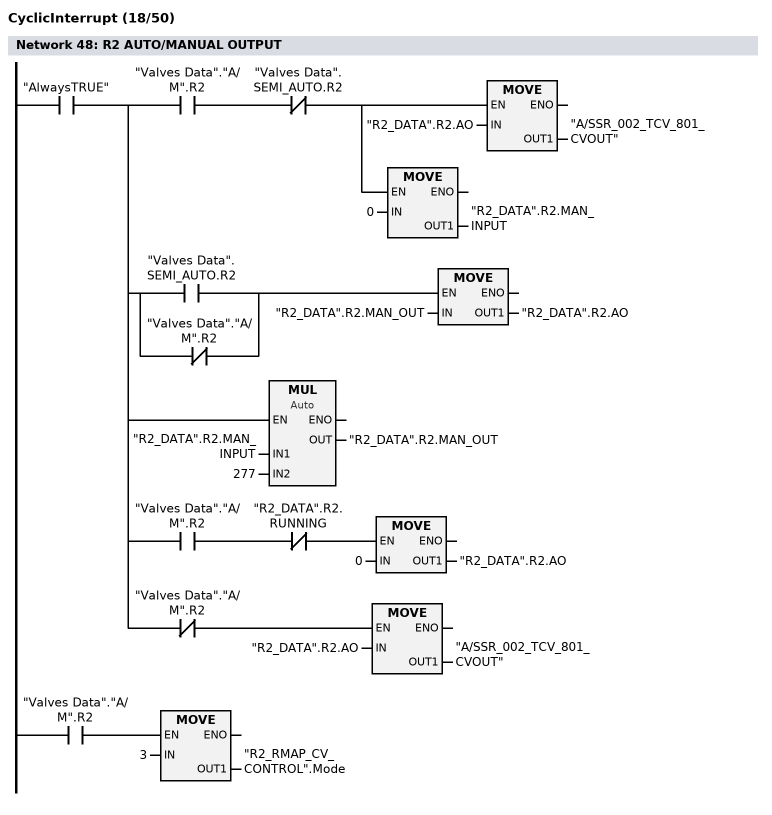
   RUNG wire#powerrail
      Contact( "AlwaysTRUE" )
      wire#w1
      Contact( "Valves Data"."A/M".R2 )
      I_Contact( "Valves Data".SEMI_AUTO.R2 )
      wire#w2
      Move(in := "R2_DATA".R2.AO, out1 => "A/SSR_002_TCV_801_CVOUT")
   END_RUNG
   RUNG wire#w2
      Move(in := 0, out1 => "R2_DATA".R2.MAN_INPUT)
   END_RUNG
   RUNG wire#w1
      Contact( "Valves Data".SEMI_AUTO.R2 )
      wire#w3
      Move(in := "R2_DATA".R2.MAN_OUT, out1 => "R2_DATA".R2.AO)
   END_RUNG
   RUNG wire#w1
      I_Contact( "Valves Data"."A/M".R2 )
   END_RUNG wire#w3
   RUNG wire#w1
      Mul(in1 := "R2_DATA".R2.MAN_INPUT, in2 := 277, out => "R2_DATA".R2.MAN_OUT)
   END_RUNG
   RUNG wire#w1
      Contact( "Valves Data"."A/M".R2 )
      I_Contact( "R2_DATA".R2.RUNNING )
      Move(in := 0, out1 => "R2_DATA".R2.AO)
   END_RUNG
   RUNG wire#w1
      I_Contact( "Valves Data"."A/M".R2 )
      Move(in := "R2_DATA".R2.AO, out1 => "A/SSR_002_TCV_801_CVOUT")
   END_RUNG
   RUNG wire#powerrail
      Contact( "Valves Data"."A/M".R2 )
      Move(in := 3, out1 => "R2_RMAP_CV_CONTROL".Mode)
   END_RUNG
   // the same network as SCL:
   IF "AlwaysTRUE" AND "Valves Data"."A/M".R2 AND NOT "Valves Data".SEMI_AUTO.R2 THEN
       "A/SSR_002_TCV_801_CVOUT" := "R2_DATA".R2.AO;
       "R2_DATA".R2.MAN_INPUT := 0;
   END_IF;
   IF "AlwaysTRUE" AND ("Valves Data".SEMI_AUTO.R2 OR NOT "Valves Data"."A/M".R2) THEN
       "R2_DATA".R2.AO := "R2_DATA".R2.MAN_OUT;
   END_IF;
   IF "AlwaysTRUE" THEN "R2_DATA".R2.MAN_OUT := "R2_DATA".R2.MAN_INPUT * 277; END_IF;
   IF "AlwaysTRUE" AND "Valves Data"."A/M".R2 AND NOT "R2_DATA".R2.RUNNING THEN "R2_DATA".R2.AO := 0; END_IF;
   IF "AlwaysTRUE" AND NOT "Valves Data"."A/M".R2 THEN "A/SSR_002_TCV_801_CVOUT" := "R2_DATA".R2.AO; END_IF;
   IF "Valves Data"."A/M".R2 THEN "R2_RMAP_CV_CONTROL".Mode := 3; END_IF;
END_REGION

REGION Network 49: R3_RAMP_CV
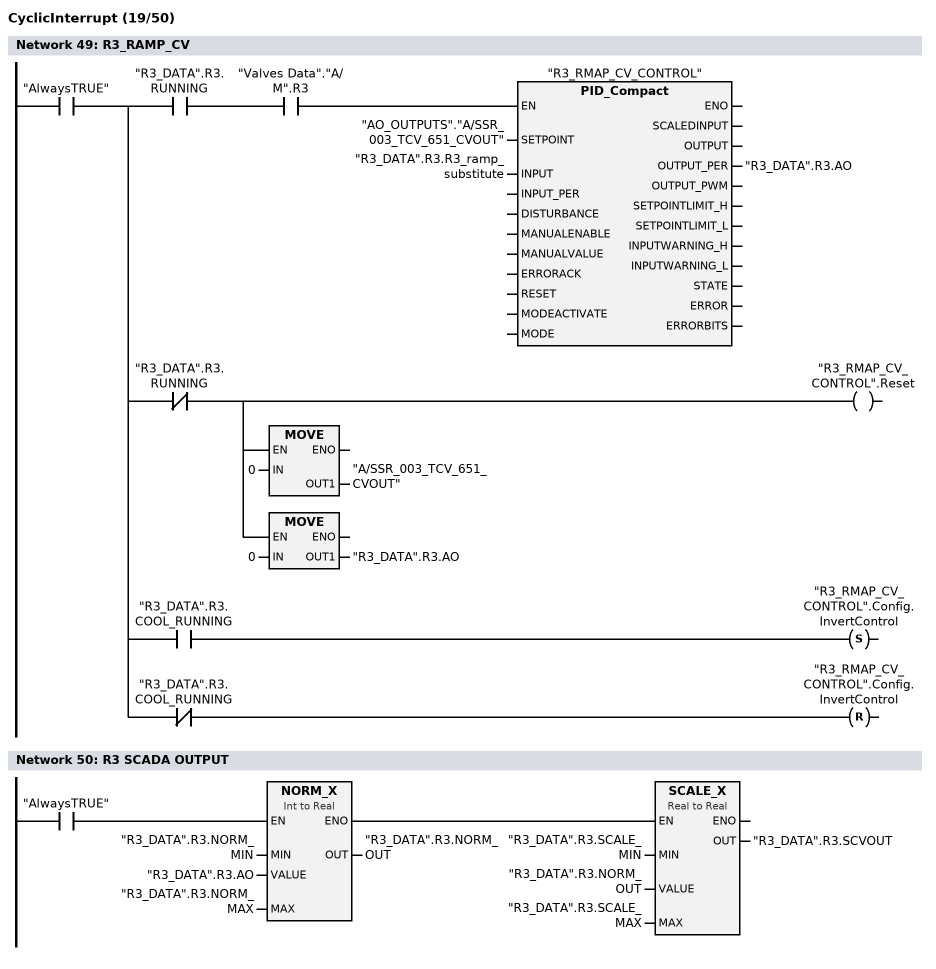
   RUNG wire#powerrail
      Contact( "AlwaysTRUE" )
      wire#w1
      Contact( "R3_DATA".R3.RUNNING )
      Contact( "Valves Data"."A/M".R3 )
      "R3_RMAP_CV_CONTROL".PID_Compact(Setpoint := "AO_OUTPUTS"."A/SSR_003_TCV_651_CVOUT", Input := "R3_DATA".R3.R3_ramp_substitute, Input_PER :=, Disturbance :=, ManualEnable :=, ManualValue :=, ErrorAck :=, Reset :=, ModeActivate :=, Mode :=, ScaledInput =>, Output =>, Output_PER => "R3_DATA".R3.AO, Output_PWM =>, SetpointLimit_H =>, SetpointLimit_L =>, InputWarning_H =>, InputWarning_L =>, State =>, Error =>, ErrorBits =>)
   END_RUNG
   RUNG wire#w1
      I_Contact( "R3_DATA".R3.RUNNING )
      wire#w2
      Coil( "R3_RMAP_CV_CONTROL".Reset )
   END_RUNG
   RUNG wire#w2
      Move(in := 0, out1 => "A/SSR_003_TCV_651_CVOUT")
   END_RUNG
   RUNG wire#w2
      Move(in := 0, out1 => "R3_DATA".R3.AO)
   END_RUNG
   RUNG wire#w1
      Contact( "R3_DATA".R3.COOL_RUNNING )
      S_Coil( "R3_RMAP_CV_CONTROL".Config.InvertControl )
   END_RUNG
   RUNG wire#w1
      I_Contact( "R3_DATA".R3.COOL_RUNNING )
      R_Coil( "R3_RMAP_CV_CONTROL".Config.InvertControl )
   END_RUNG
   // the same network as SCL:
   #_w1 := "AlwaysTRUE";
   IF "AlwaysTRUE" AND "R3_DATA".R3.RUNNING AND "Valves Data"."A/M".R3 THEN
       "R3_RMAP_CV_CONTROL"(Setpoint := "AO_OUTPUTS"."A/SSR_003_TCV_651_CVOUT",   // PID_Compact
                            Input := "R3_DATA".R3.R3_ramp_substitute,
                            Output_PER => "R3_DATA".R3.AO);
   END_IF;
   "R3_RMAP_CV_CONTROL".Reset := #_w1 AND NOT "R3_DATA".R3.RUNNING;
   IF "R3_RMAP_CV_CONTROL".Reset THEN
       "A/SSR_003_TCV_651_CVOUT" := 0;
       "R3_DATA".R3.AO := 0;
   END_IF;
   IF #_w1 AND "R3_DATA".R3.COOL_RUNNING THEN "R3_RMAP_CV_CONTROL".Config.InvertControl := TRUE; END_IF;
   IF #_w1 AND NOT "R3_DATA".R3.COOL_RUNNING THEN "R3_RMAP_CV_CONTROL".Config.InvertControl := FALSE; END_IF;
END_REGION

REGION Network 50: R3 SCADA OUTPUT
   RUNG wire#powerrail
      Contact( "AlwaysTRUE" )
      { S7_Templates := "[SrcType := Int, DestType := Real]" } Normalize(min := "R3_DATA".R3.NORM_MIN, value := "R3_DATA".R3.AO, max := "R3_DATA".R3.NORM_MAX, out => "R3_DATA".R3.NORM_OUT)
      { S7_Templates := "[SrcType := Real, DestType := Real]" } Scale(min := "R3_DATA".R3.SCALE_MIN, value := "R3_DATA".R3.NORM_OUT, max := "R3_DATA".R3.SCALE_MAX, out => "R3_DATA".R3.SCVOUT)
   END_RUNG
   // the same network as SCL:
   IF "AlwaysTRUE" THEN
       "R3_DATA".R3.NORM_OUT := NORM_X(MIN := "R3_DATA".R3.NORM_MIN, VALUE := "R3_DATA".R3.AO, MAX := "R3_DATA".R3.NORM_MAX);
       "R3_DATA".R3.SCVOUT := SCALE_X(MIN := "R3_DATA".R3.SCALE_MIN, VALUE := "R3_DATA".R3.NORM_OUT, MAX := "R3_DATA".R3.SCALE_MAX);
   END_IF;
END_REGION

REGION Network 51: R3 AUTO/MANUAL OUTPUT
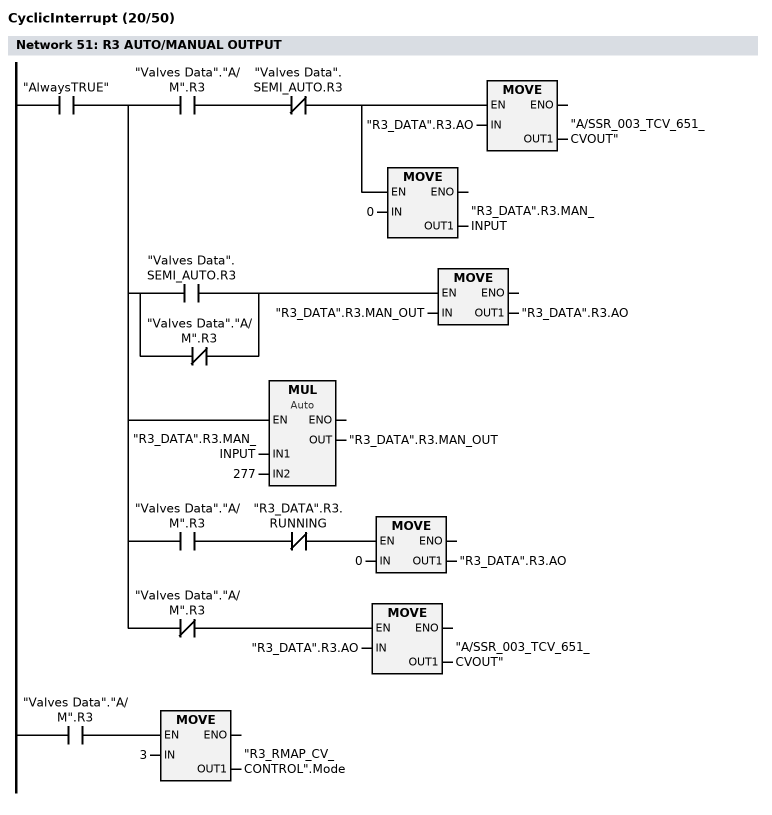
   RUNG wire#powerrail
      Contact( "AlwaysTRUE" )
      wire#w1
      Contact( "Valves Data"."A/M".R3 )
      I_Contact( "Valves Data".SEMI_AUTO.R3 )
      wire#w2
      Move(in := "R3_DATA".R3.AO, out1 => "A/SSR_003_TCV_651_CVOUT")
   END_RUNG
   RUNG wire#w2
      Move(in := 0, out1 => "R3_DATA".R3.MAN_INPUT)
   END_RUNG
   RUNG wire#w1
      Contact( "Valves Data".SEMI_AUTO.R3 )
      wire#w3
      Move(in := "R3_DATA".R3.MAN_OUT, out1 => "R3_DATA".R3.AO)
   END_RUNG
   RUNG wire#w1
      I_Contact( "Valves Data"."A/M".R3 )
   END_RUNG wire#w3
   RUNG wire#w1
      Mul(in1 := "R3_DATA".R3.MAN_INPUT, in2 := 277, out => "R3_DATA".R3.MAN_OUT)
   END_RUNG
   RUNG wire#w1
      Contact( "Valves Data"."A/M".R3 )
      I_Contact( "R3_DATA".R3.RUNNING )
      Move(in := 0, out1 => "R3_DATA".R3.AO)
   END_RUNG
   RUNG wire#w1
      I_Contact( "Valves Data"."A/M".R3 )
      Move(in := "R3_DATA".R3.AO, out1 => "A/SSR_003_TCV_651_CVOUT")
   END_RUNG
   RUNG wire#powerrail
      Contact( "Valves Data"."A/M".R3 )
      Move(in := 3, out1 => "R3_RMAP_CV_CONTROL".Mode)
   END_RUNG
   // the same network as SCL:
   IF "AlwaysTRUE" AND "Valves Data"."A/M".R3 AND NOT "Valves Data".SEMI_AUTO.R3 THEN
       "A/SSR_003_TCV_651_CVOUT" := "R3_DATA".R3.AO;
       "R3_DATA".R3.MAN_INPUT := 0;
   END_IF;
   IF "AlwaysTRUE" AND ("Valves Data".SEMI_AUTO.R3 OR NOT "Valves Data"."A/M".R3) THEN
       "R3_DATA".R3.AO := "R3_DATA".R3.MAN_OUT;
   END_IF;
   IF "AlwaysTRUE" THEN "R3_DATA".R3.MAN_OUT := "R3_DATA".R3.MAN_INPUT * 277; END_IF;
   IF "AlwaysTRUE" AND "Valves Data"."A/M".R3 AND NOT "R3_DATA".R3.RUNNING THEN "R3_DATA".R3.AO := 0; END_IF;
   IF "AlwaysTRUE" AND NOT "Valves Data"."A/M".R3 THEN "A/SSR_003_TCV_651_CVOUT" := "R3_DATA".R3.AO; END_IF;
   IF "Valves Data"."A/M".R3 THEN "R3_RMAP_CV_CONTROL".Mode := 3; END_IF;
END_REGION

REGION Network 52: R4_RAMP_CV
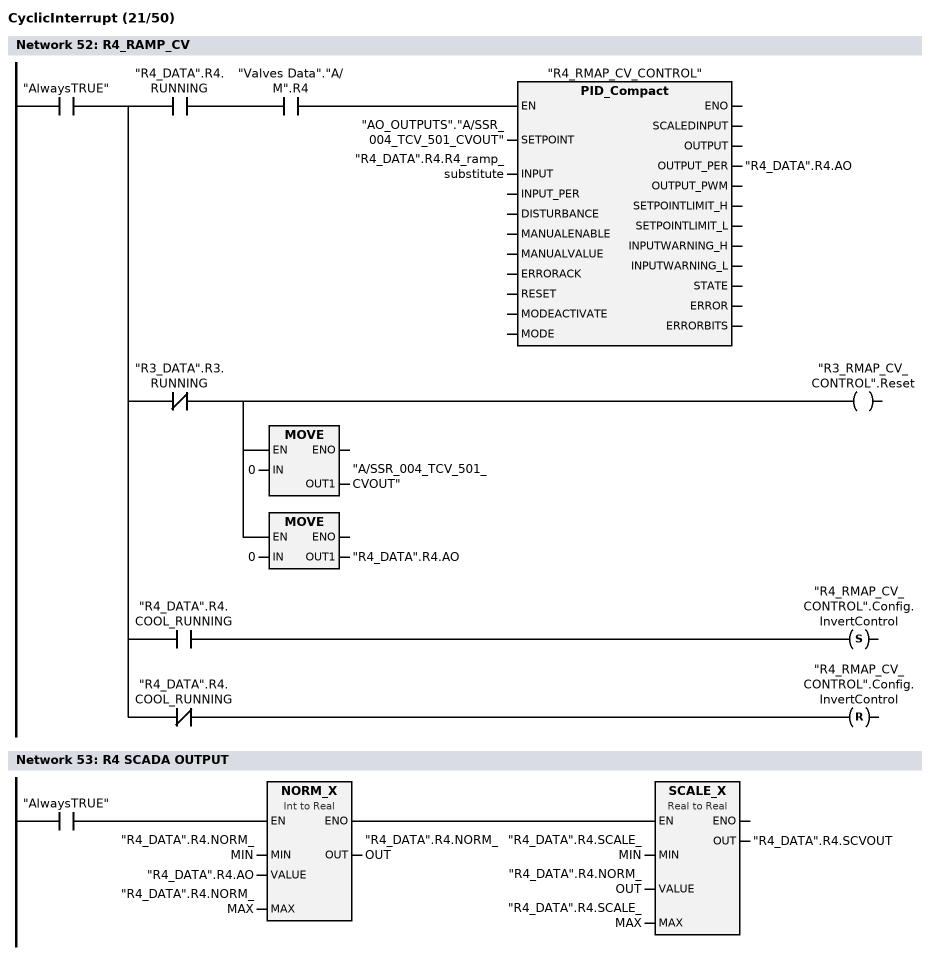
   RUNG wire#powerrail
      Contact( "AlwaysTRUE" )
      wire#w1
      Contact( "R4_DATA".R4.RUNNING )
      Contact( "Valves Data"."A/M".R4 )
      "R4_RMAP_CV_CONTROL".PID_Compact(Setpoint := "AO_OUTPUTS"."A/SSR_004_TCV_501_CVOUT", Input := "R4_DATA".R4.R4_ramp_substitute, Input_PER :=, Disturbance :=, ManualEnable :=, ManualValue :=, ErrorAck :=, Reset :=, ModeActivate :=, Mode :=, ScaledInput =>, Output =>, Output_PER => "R4_DATA".R4.AO, Output_PWM =>, SetpointLimit_H =>, SetpointLimit_L =>, InputWarning_H =>, InputWarning_L =>, State =>, Error =>, ErrorBits =>)
   END_RUNG
   RUNG wire#w1
      I_Contact( "R3_DATA".R3.RUNNING )
      wire#w2
      Coil( "R3_RMAP_CV_CONTROL".Reset )
   END_RUNG
   RUNG wire#w2
      Move(in := 0, out1 => "A/SSR_004_TCV_501_CVOUT")
   END_RUNG
   RUNG wire#w2
      Move(in := 0, out1 => "R4_DATA".R4.AO)
   END_RUNG
   RUNG wire#w1
      Contact( "R4_DATA".R4.COOL_RUNNING )
      S_Coil( "R4_RMAP_CV_CONTROL".Config.InvertControl )
   END_RUNG
   RUNG wire#w1
      I_Contact( "R4_DATA".R4.COOL_RUNNING )
      R_Coil( "R4_RMAP_CV_CONTROL".Config.InvertControl )
   END_RUNG
   // the same network as SCL:
   #_w1 := "AlwaysTRUE";
   IF "AlwaysTRUE" AND "R4_DATA".R4.RUNNING AND "Valves Data"."A/M".R4 THEN
       "R4_RMAP_CV_CONTROL"(Setpoint := "AO_OUTPUTS"."A/SSR_004_TCV_501_CVOUT",   // PID_Compact
                            Input := "R4_DATA".R4.R4_ramp_substitute,
                            Output_PER => "R4_DATA".R4.AO);
   END_IF;
   "R3_RMAP_CV_CONTROL".Reset := #_w1 AND NOT "R3_DATA".R3.RUNNING;
   IF "R3_RMAP_CV_CONTROL".Reset THEN
       "A/SSR_004_TCV_501_CVOUT" := 0;
       "R4_DATA".R4.AO := 0;
   END_IF;
   IF #_w1 AND "R4_DATA".R4.COOL_RUNNING THEN "R4_RMAP_CV_CONTROL".Config.InvertControl := TRUE; END_IF;
   IF #_w1 AND NOT "R4_DATA".R4.COOL_RUNNING THEN "R4_RMAP_CV_CONTROL".Config.InvertControl := FALSE; END_IF;
END_REGION

REGION Network 53: R4 SCADA OUTPUT
   RUNG wire#powerrail
      Contact( "AlwaysTRUE" )
      { S7_Templates := "[SrcType := Int, DestType := Real]" } Normalize(min := "R4_DATA".R4.NORM_MIN, value := "R4_DATA".R4.AO, max := "R4_DATA".R4.NORM_MAX, out => "R4_DATA".R4.NORM_OUT)
      { S7_Templates := "[SrcType := Real, DestType := Real]" } Scale(min := "R4_DATA".R4.SCALE_MIN, value := "R4_DATA".R4.NORM_OUT, max := "R4_DATA".R4.SCALE_MAX, out => "R4_DATA".R4.SCVOUT)
   END_RUNG
   // the same network as SCL:
   IF "AlwaysTRUE" THEN
       "R4_DATA".R4.NORM_OUT := NORM_X(MIN := "R4_DATA".R4.NORM_MIN, VALUE := "R4_DATA".R4.AO, MAX := "R4_DATA".R4.NORM_MAX);
       "R4_DATA".R4.SCVOUT := SCALE_X(MIN := "R4_DATA".R4.SCALE_MIN, VALUE := "R4_DATA".R4.NORM_OUT, MAX := "R4_DATA".R4.SCALE_MAX);
   END_IF;
END_REGION

REGION Network 54: R4 AUTO/MANUAL OUTPUT
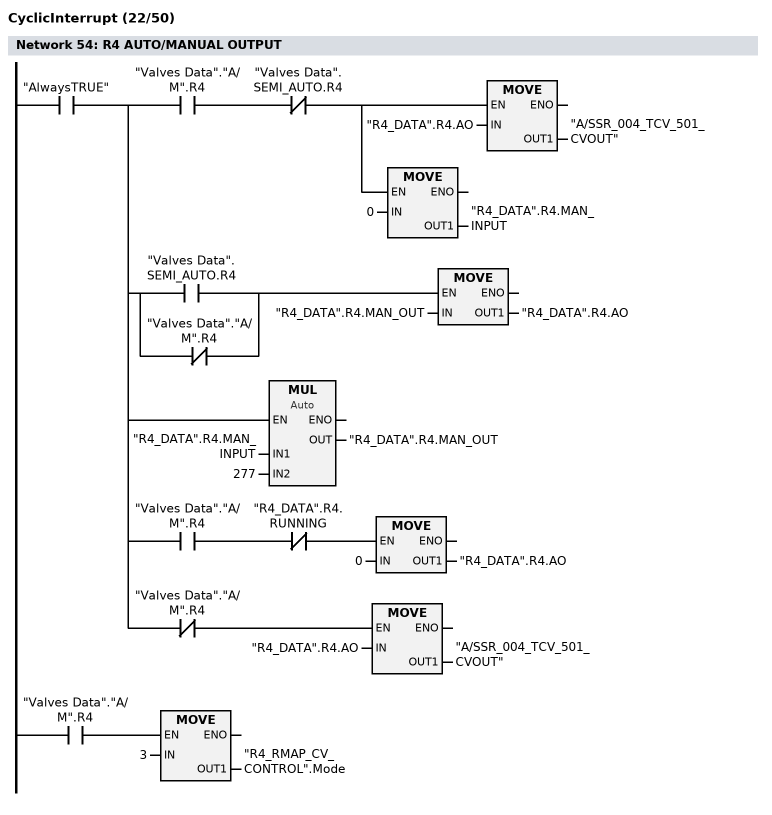
   RUNG wire#powerrail
      Contact( "AlwaysTRUE" )
      wire#w1
      Contact( "Valves Data"."A/M".R4 )
      I_Contact( "Valves Data".SEMI_AUTO.R4 )
      wire#w2
      Move(in := "R4_DATA".R4.AO, out1 => "A/SSR_004_TCV_501_CVOUT")
   END_RUNG
   RUNG wire#w2
      Move(in := 0, out1 => "R4_DATA".R4.MAN_INPUT)
   END_RUNG
   RUNG wire#w1
      Contact( "Valves Data".SEMI_AUTO.R4 )
      wire#w3
      Move(in := "R4_DATA".R4.MAN_OUT, out1 => "R4_DATA".R4.AO)
   END_RUNG
   RUNG wire#w1
      I_Contact( "Valves Data"."A/M".R4 )
   END_RUNG wire#w3
   RUNG wire#w1
      Mul(in1 := "R4_DATA".R4.MAN_INPUT, in2 := 277, out => "R4_DATA".R4.MAN_OUT)
   END_RUNG
   RUNG wire#w1
      Contact( "Valves Data"."A/M".R4 )
      I_Contact( "R4_DATA".R4.RUNNING )
      Move(in := 0, out1 => "R4_DATA".R4.AO)
   END_RUNG
   RUNG wire#w1
      I_Contact( "Valves Data"."A/M".R4 )
      Move(in := "R4_DATA".R4.AO, out1 => "A/SSR_004_TCV_501_CVOUT")
   END_RUNG
   RUNG wire#powerrail
      Contact( "Valves Data"."A/M".R4 )
      Move(in := 3, out1 => "R4_RMAP_CV_CONTROL".Mode)
   END_RUNG
   // the same network as SCL:
   IF "AlwaysTRUE" AND "Valves Data"."A/M".R4 AND NOT "Valves Data".SEMI_AUTO.R4 THEN
       "A/SSR_004_TCV_501_CVOUT" := "R4_DATA".R4.AO;
       "R4_DATA".R4.MAN_INPUT := 0;
   END_IF;
   IF "AlwaysTRUE" AND ("Valves Data".SEMI_AUTO.R4 OR NOT "Valves Data"."A/M".R4) THEN
       "R4_DATA".R4.AO := "R4_DATA".R4.MAN_OUT;
   END_IF;
   IF "AlwaysTRUE" THEN "R4_DATA".R4.MAN_OUT := "R4_DATA".R4.MAN_INPUT * 277; END_IF;
   IF "AlwaysTRUE" AND "Valves Data"."A/M".R4 AND NOT "R4_DATA".R4.RUNNING THEN "R4_DATA".R4.AO := 0; END_IF;
   IF "AlwaysTRUE" AND NOT "Valves Data"."A/M".R4 THEN "A/SSR_004_TCV_501_CVOUT" := "R4_DATA".R4.AO; END_IF;
   IF "Valves Data"."A/M".R4 THEN "R4_RMAP_CV_CONTROL".Mode := 3; END_IF;
END_REGION

REGION Network 55: R5_RAMP_CV
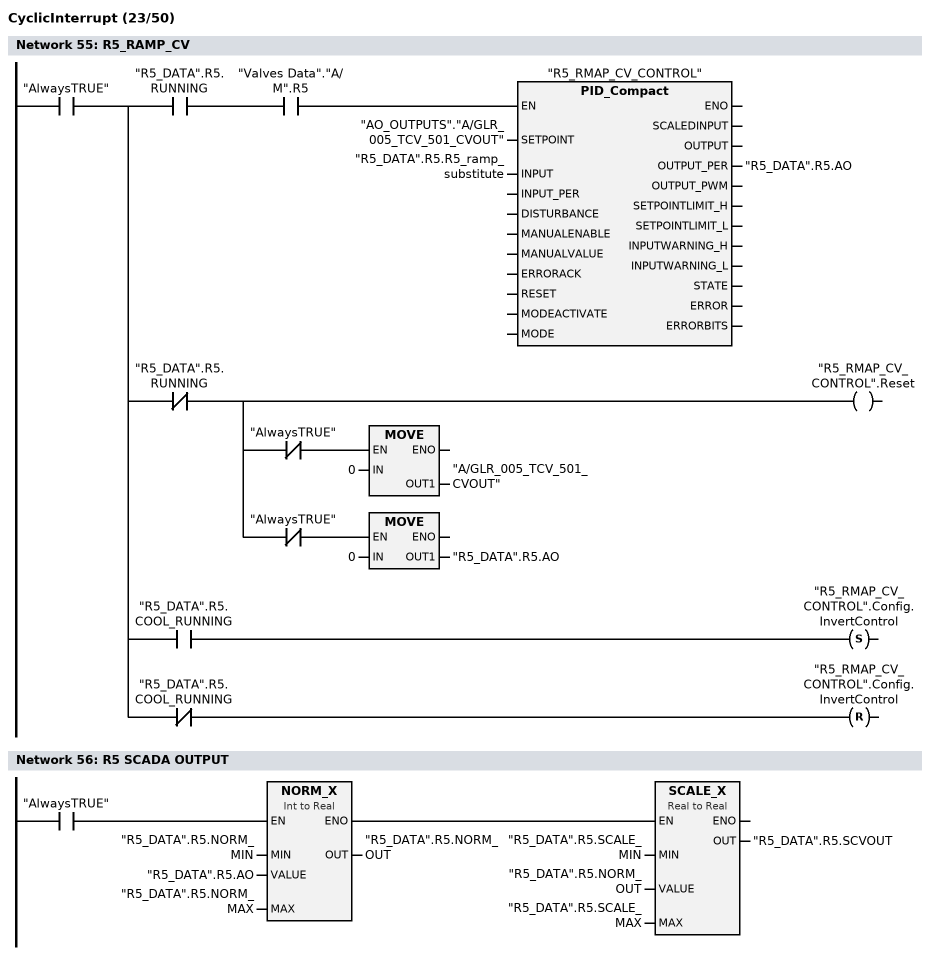
   RUNG wire#powerrail
      Contact( "AlwaysTRUE" )
      wire#w1
      Contact( "R5_DATA".R5.RUNNING )
      Contact( "Valves Data"."A/M".R5 )
      "R5_RMAP_CV_CONTROL".PID_Compact(Setpoint := "AO_OUTPUTS"."A/GLR_005_TCV_501_CVOUT", Input := "R5_DATA".R5.R5_ramp_substitute, Input_PER :=, Disturbance :=, ManualEnable :=, ManualValue :=, ErrorAck :=, Reset :=, ModeActivate :=, Mode :=, ScaledInput =>, Output =>, Output_PER => "R5_DATA".R5.AO, Output_PWM =>, SetpointLimit_H =>, SetpointLimit_L =>, InputWarning_H =>, InputWarning_L =>, State =>, Error =>, ErrorBits =>)
   END_RUNG
   RUNG wire#w1
      I_Contact( "R5_DATA".R5.RUNNING )
      wire#w2
      Coil( "R5_RMAP_CV_CONTROL".Reset )
   END_RUNG
   RUNG wire#w2
      I_Contact( "AlwaysTRUE" )
      Move(in := 0, out1 => "A/GLR_005_TCV_501_CVOUT")
   END_RUNG
   RUNG wire#w2
      I_Contact( "AlwaysTRUE" )
      Move(in := 0, out1 => "R5_DATA".R5.AO)
   END_RUNG
   RUNG wire#w1
      Contact( "R5_DATA".R5.COOL_RUNNING )
      S_Coil( "R5_RMAP_CV_CONTROL".Config.InvertControl )
   END_RUNG
   RUNG wire#w1
      I_Contact( "R5_DATA".R5.COOL_RUNNING )
      R_Coil( "R5_RMAP_CV_CONTROL".Config.InvertControl )
   END_RUNG
   // the same network as SCL:
   #_w1 := "AlwaysTRUE";
   IF "AlwaysTRUE" AND "R5_DATA".R5.RUNNING AND "Valves Data"."A/M".R5 THEN
       "R5_RMAP_CV_CONTROL"(Setpoint := "AO_OUTPUTS"."A/GLR_005_TCV_501_CVOUT",   // PID_Compact
                            Input := "R5_DATA".R5.R5_ramp_substitute,
                            Output_PER => "R5_DATA".R5.AO);
   END_IF;
   "R5_RMAP_CV_CONTROL".Reset := #_w1 AND NOT "R5_DATA".R5.RUNNING;
   IF "R5_RMAP_CV_CONTROL".Reset AND NOT "AlwaysTRUE" THEN
       "A/GLR_005_TCV_501_CVOUT" := 0;
       "R5_DATA".R5.AO := 0;
   END_IF;
   IF #_w1 AND "R5_DATA".R5.COOL_RUNNING THEN "R5_RMAP_CV_CONTROL".Config.InvertControl := TRUE; END_IF;
   IF #_w1 AND NOT "R5_DATA".R5.COOL_RUNNING THEN "R5_RMAP_CV_CONTROL".Config.InvertControl := FALSE; END_IF;
END_REGION

REGION Network 56: R5 SCADA OUTPUT
   RUNG wire#powerrail
      Contact( "AlwaysTRUE" )
      { S7_Templates := "[SrcType := Int, DestType := Real]" } Normalize(min := "R5_DATA".R5.NORM_MIN, value := "R5_DATA".R5.AO, max := "R5_DATA".R5.NORM_MAX, out => "R5_DATA".R5.NORM_OUT)
      { S7_Templates := "[SrcType := Real, DestType := Real]" } Scale(min := "R5_DATA".R5.SCALE_MIN, value := "R5_DATA".R5.NORM_OUT, max := "R5_DATA".R5.SCALE_MAX, out => "R5_DATA".R5.SCVOUT)
   END_RUNG
   // the same network as SCL:
   IF "AlwaysTRUE" THEN
       "R5_DATA".R5.NORM_OUT := NORM_X(MIN := "R5_DATA".R5.NORM_MIN, VALUE := "R5_DATA".R5.AO, MAX := "R5_DATA".R5.NORM_MAX);
       "R5_DATA".R5.SCVOUT := SCALE_X(MIN := "R5_DATA".R5.SCALE_MIN, VALUE := "R5_DATA".R5.NORM_OUT, MAX := "R5_DATA".R5.SCALE_MAX);
   END_IF;
END_REGION

REGION Network 57: R5 AUTO/MANUAL OUTPUT
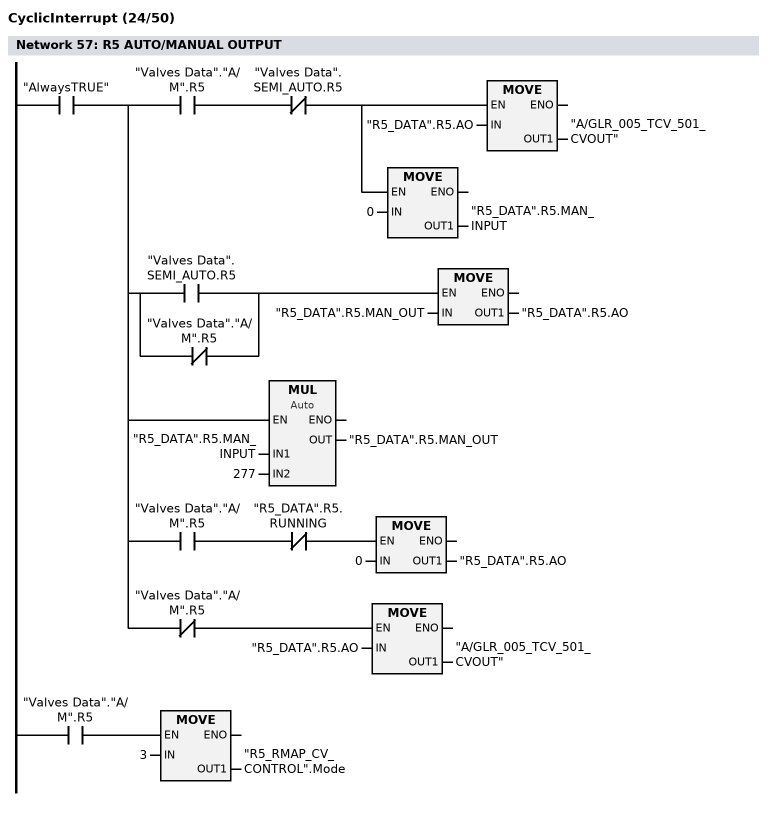
   RUNG wire#powerrail
      Contact( "AlwaysTRUE" )
      wire#w1
      Contact( "Valves Data"."A/M".R5 )
      I_Contact( "Valves Data".SEMI_AUTO.R5 )
      wire#w2
      Move(in := "R5_DATA".R5.AO, out1 => "A/GLR_005_TCV_501_CVOUT")
   END_RUNG
   RUNG wire#w2
      Move(in := 0, out1 => "R5_DATA".R5.MAN_INPUT)
   END_RUNG
   RUNG wire#w1
      Contact( "Valves Data".SEMI_AUTO.R5 )
      wire#w3
      Move(in := "R5_DATA".R5.MAN_OUT, out1 => "R5_DATA".R5.AO)
   END_RUNG
   RUNG wire#w1
      I_Contact( "Valves Data"."A/M".R5 )
   END_RUNG wire#w3
   RUNG wire#w1
      Mul(in1 := "R5_DATA".R5.MAN_INPUT, in2 := 277, out => "R5_DATA".R5.MAN_OUT)
   END_RUNG
   RUNG wire#w1
      Contact( "Valves Data"."A/M".R5 )
      I_Contact( "R5_DATA".R5.RUNNING )
      Move(in := 0, out1 => "R5_DATA".R5.AO)
   END_RUNG
   RUNG wire#w1
      I_Contact( "Valves Data"."A/M".R5 )
      Move(in := "R5_DATA".R5.AO, out1 => "A/GLR_005_TCV_501_CVOUT")
   END_RUNG
   RUNG wire#powerrail
      Contact( "Valves Data"."A/M".R5 )
      Move(in := 3, out1 => "R5_RMAP_CV_CONTROL".Mode)
   END_RUNG
   // the same network as SCL:
   IF "AlwaysTRUE" AND "Valves Data"."A/M".R5 AND NOT "Valves Data".SEMI_AUTO.R5 THEN
       "A/GLR_005_TCV_501_CVOUT" := "R5_DATA".R5.AO;
       "R5_DATA".R5.MAN_INPUT := 0;
   END_IF;
   IF "AlwaysTRUE" AND ("Valves Data".SEMI_AUTO.R5 OR NOT "Valves Data"."A/M".R5) THEN
       "R5_DATA".R5.AO := "R5_DATA".R5.MAN_OUT;
   END_IF;
   IF "AlwaysTRUE" THEN "R5_DATA".R5.MAN_OUT := "R5_DATA".R5.MAN_INPUT * 277; END_IF;
   IF "AlwaysTRUE" AND "Valves Data"."A/M".R5 AND NOT "R5_DATA".R5.RUNNING THEN "R5_DATA".R5.AO := 0; END_IF;
   IF "AlwaysTRUE" AND NOT "Valves Data"."A/M".R5 THEN "A/GLR_005_TCV_501_CVOUT" := "R5_DATA".R5.AO; END_IF;
   IF "Valves Data"."A/M".R5 THEN "R5_RMAP_CV_CONTROL".Mode := 3; END_IF;
END_REGION

REGION Network 58: R6_RAMP_CV
